(* IEC 61131-3 sources: Aqueous_Solutions/docs-authority/plc (part 3) *)

(* ---- PLC-HEAT.st ---- *)
(* AQS-CTL-004 X-CTL-04: control program source, generated by flow_graph/control/plc_programs.py *)
(* Basis: AQS-CTL-001 INSTRUMENT_INDEX.csv, AQS-CTL-002 control architecture, graph set-points. *)
(* PLC-HEAT: CPU single; IO counts AI 24 AO 0 DI 0 DO 0 (modules per AQS-CTL-002, 16-channel, 20 % spare) *)
PROGRAM PLC_HEAT_CTRL
VAR
  (* 100 ms cyclic task per AQS-CTL-002 *)
  DRY_COOLERPT-01_PV : REAL ;  (* no design pressure on the graph )
  DRY_COOLERTE-01_PV : REAL ;  (* band by service )
  Q1_APT-01_PV : REAL ;  (* no design pressure on the graph )
  Q1_ATE-01_PV : REAL ;  (* band by service )
  Q1_BPT-01_PV : REAL ;  (* no design pressure on the graph )
  Q1_BTE-01_PV : REAL ;  (* band by service )
  Q2_APT-01_PV : REAL ;  (* no design pressure on the graph )
  Q2_ATE-01_PV : REAL ;  (* band by service )
  Q2_BPT-01_PV : REAL ;  (* no design pressure on the graph )
  Q2_BTE-01_PV : REAL ;  (* band by service )
  Q3_APT-01_PV : REAL ;  (* no design pressure on the graph )
  Q3_ATE-01_PV : REAL ;  (* band by service )
  Q3_BPT-01_PV : REAL ;  (* no design pressure on the graph )
  Q3_BTE-01_PV : REAL ;  (* band by service )
  Q4_APT-01_PV : REAL ;  (* no design pressure on the graph )
  Q4_ATE-01_PV : REAL ;  (* band by service )
  Q4_BPT-01_PV : REAL ;  (* no design pressure on the graph )
  Q4_BTE-01_PV : REAL ;  (* band by service )
  ADS_CHILLTE-01_PV : REAL ;  (* drive water in: IA-Q4-ADS 5.0 kW Q4 65 C )
  ADS_CHILLTE-02_PV : REAL ;  (* chilled water out: IA-ADS-CHW 2.25 kW at 12 C )
  MAU_HXTE-01_PV : REAL ;  (* Q4 coil: IA-Q4-MAU 12 kW Q4 water 65/45 C (winter design) )
  Q4_BUSTE-01_PV : REAL ;  (* Q4 hot-water bus supply (IA-Q4-ADS/IA-Q4-MAU 65 C design) )
  Q4_BUSPT-01_PV : REAL ;  (* hot-water bus; no design pressure on the graph )
  RAD_PANELTE-01_PV : REAL ;  (* radiator loop outlet temperature watch; rejection performance against the A-M-39 )
END_VAR

  (* PRESSURE monitoring block - indication, no set-point invented )
  FB_AI_DRY_COOLERPT-01( PV := DRY_COOLERPT-01_PV );
  DRY_COOLERPT-01_ALARM_HI := 9.0 ;  (* 90 % of span, registered LSH convention )

  (* TEMPERATURE monitoring block - indication, no set-point invented )
  FB_AI_DRY_COOLERTE-01( PV := DRY_COOLERTE-01_PV );
  DRY_COOLERTE-01_ALARM_HI := 135.0 ;  (* 90 % of span, registered LSH convention )

  (* PRESSURE monitoring block - indication, no set-point invented )
  FB_AI_Q1_APT-01( PV := Q1_APT-01_PV );
  Q1_APT-01_ALARM_HI := 9.0 ;  (* 90 % of span, registered LSH convention )

  (* TEMPERATURE monitoring block - indication, no set-point invented )
  FB_AI_Q1_ATE-01( PV := Q1_ATE-01_PV );
  Q1_ATE-01_ALARM_HI := 135.0 ;  (* 90 % of span, registered LSH convention )

  (* PRESSURE monitoring block - indication, no set-point invented )
  FB_AI_Q1_BPT-01( PV := Q1_BPT-01_PV );
  Q1_BPT-01_ALARM_HI := 9.0 ;  (* 90 % of span, registered LSH convention )

  (* TEMPERATURE monitoring block - indication, no set-point invented )
  FB_AI_Q1_BTE-01( PV := Q1_BTE-01_PV );
  Q1_BTE-01_ALARM_HI := 135.0 ;  (* 90 % of span, registered LSH convention )

  (* PRESSURE monitoring block - indication, no set-point invented )
  FB_AI_Q2_APT-01( PV := Q2_APT-01_PV );
  Q2_APT-01_ALARM_HI := 9.0 ;  (* 90 % of span, registered LSH convention )

  (* TEMPERATURE monitoring block - indication, no set-point invented )
  FB_AI_Q2_ATE-01( PV := Q2_ATE-01_PV );
  Q2_ATE-01_ALARM_HI := 135.0 ;  (* 90 % of span, registered LSH convention )

  (* PRESSURE monitoring block - indication, no set-point invented )
  FB_AI_Q2_BPT-01( PV := Q2_BPT-01_PV );
  Q2_BPT-01_ALARM_HI := 9.0 ;  (* 90 % of span, registered LSH convention )

  (* TEMPERATURE monitoring block - indication, no set-point invented )
  FB_AI_Q2_BTE-01( PV := Q2_BTE-01_PV );
  Q2_BTE-01_ALARM_HI := 135.0 ;  (* 90 % of span, registered LSH convention )

  (* PRESSURE monitoring block - indication, no set-point invented )
  FB_AI_Q3_APT-01( PV := Q3_APT-01_PV );
  Q3_APT-01_ALARM_HI := 9.0 ;  (* 90 % of span, registered LSH convention )

  (* TEMPERATURE monitoring block - indication, no set-point invented )
  FB_AI_Q3_ATE-01( PV := Q3_ATE-01_PV );
  Q3_ATE-01_ALARM_HI := 135.0 ;  (* 90 % of span, registered LSH convention )

  (* PRESSURE monitoring block - indication, no set-point invented )
  FB_AI_Q3_BPT-01( PV := Q3_BPT-01_PV );
  Q3_BPT-01_ALARM_HI := 9.0 ;  (* 90 % of span, registered LSH convention )

  (* TEMPERATURE monitoring block - indication, no set-point invented )
  FB_AI_Q3_BTE-01( PV := Q3_BTE-01_PV );
  Q3_BTE-01_ALARM_HI := 135.0 ;  (* 90 % of span, registered LSH convention )

  (* PRESSURE monitoring block - indication, no set-point invented )
  FB_AI_Q4_APT-01( PV := Q4_APT-01_PV );
  Q4_APT-01_ALARM_HI := 9.0 ;  (* 90 % of span, registered LSH convention )

  (* TEMPERATURE monitoring block - indication, no set-point invented )
  FB_AI_Q4_ATE-01( PV := Q4_ATE-01_PV );
  Q4_ATE-01_ALARM_HI := 135.0 ;  (* 90 % of span, registered LSH convention )

  (* PRESSURE monitoring block - indication, no set-point invented )
  FB_AI_Q4_BPT-01( PV := Q4_BPT-01_PV );
  Q4_BPT-01_ALARM_HI := 9.0 ;  (* 90 % of span, registered LSH convention )

  (* TEMPERATURE monitoring block - indication, no set-point invented )
  FB_AI_Q4_BTE-01( PV := Q4_BTE-01_PV );
  Q4_BTE-01_ALARM_HI := 135.0 ;  (* 90 % of span, registered LSH convention )

  (* TEMPERATURE monitoring block - indication, no set-point invented )
  FB_AI_ADS_CHILLTE-01( PV := ADS_CHILLTE-01_PV );
  ADS_CHILLTE-01_ALARM_HI := 90.0 ;  (* 90 % of span, registered LSH convention )

  (* TEMPERATURE monitoring block - indication, no set-point invented )
  FB_AI_ADS_CHILLTE-02( PV := ADS_CHILLTE-02_PV );
  ADS_CHILLTE-02_ALARM_HI := 36.0 ;  (* 90 % of span, registered LSH convention )

  (* TEMPERATURE monitoring block - indication, no set-point invented )
  FB_AI_MAU_HXTE-01( PV := MAU_HXTE-01_PV );
  MAU_HXTE-01_ALARM_HI := 90.0 ;  (* 90 % of span, registered LSH convention )

  (* TEMPERATURE monitoring block - indication, no set-point invented )
  FB_AI_Q4_BUSTE-01( PV := Q4_BUSTE-01_PV );
  Q4_BUSTE-01_ALARM_HI := 90.0 ;  (* 90 % of span, registered LSH convention )

  (* PRESSURE monitoring block - indication, no set-point invented )
  FB_AI_Q4_BUSPT-01( PV := Q4_BUSPT-01_PV );
  Q4_BUSPT-01_ALARM_HI := 9.0 ;  (* 90 % of span, registered LSH convention )

  (* TEMPERATURE monitoring block - indication, no set-point invented )
  FB_AI_RAD_PANELTE-01( PV := RAD_PANELTE-01_PV );
  RAD_PANELTE-01_ALARM_HI := 135.0 ;  (* 90 % of span, registered LSH convention )

END_PROGRAM

(* ---- PLC-MEOH.st ---- *)
(* AQS-CTL-004 X-CTL-04: control program source, generated by flow_graph/control/plc_programs.py *)
(* Basis: AQS-CTL-001 INSTRUMENT_INDEX.csv, AQS-CTL-002 control architecture, graph set-points. *)
(* PLC-MEOH: CPU single; IO counts AI 33 AO 0 DI 51 DO 12 (modules per AQS-CTL-002, 16-channel, 20 % spare) *)
PROGRAM PLC_MEOH_CTRL
VAR
  (* 100 ms cyclic task per AQS-CTL-002 *)
  MET_SYNFT-01_PV : REAL ;  (* DL_MET_TO_FEED normal 0.00 L/h )
  MET_SYNPT-01_PV : REAL ;  (* no design pressure on the graph )
  MET_SYNTE-01_PV : REAL ;  (* band by service )
  MEOH_FERMFT-01_PV : REAL ;  (* S77 normal 0.00 L/h )
  MEOH_FERMPT-01_PV : REAL ;  (* no design pressure on the graph )
  MEOH_FERMTE-01_PV : REAL ;  (* design T 35 C )
  MEOH_FCFT-01_PV : REAL ;  (* S81 normal 0.30 L/h )
  MEOH_FCFT-02_PV : REAL ;  (* S82 normal 0.36 L/h )
  MEOH_FCFT-03_PV : REAL ;  (* IA-FC-EXH normal 0.00 L/h )
  MEOH_FCLT-01_PV : REAL ;  (* A-M-182 liquid height )
  MEOH_FCPT-01_PV : REAL ;  (* no design pressure on the graph )
  MEOH_FCTE-01_PV : REAL ;  (* band by service )
  MEOH_SYNTHFT-01_PV : REAL ;  (* IA-ESS-MEOH-CHG normal 0.00 L/h )
  MEOH_SYNTHFT-02_PV : REAL ;  (* S75 normal 1.47 L/h )
  MEOH_SYNTHFT-03_PV : REAL ;  (* MEOH_TO_OLEFIN normal 0.00 L/h )
  MEOH_SYNTHFT-04_PV : REAL ;  (* IA-MEOH-H2O normal 0.82 L/h )
  MEOH_SYNTHFT-05_PV : REAL ;  (* IA-MEOH-CH3SH normal 0.00 L/h )
  MEOH_SYNTHPT-01_PV : REAL ;  (* no design pressure on the graph )
  MEOH_SYNTHTE-01_PV : REAL ;  (* design T 250 C )
  MEOH_CONDLT-01_PV : REAL ;  (* A-M-182 liquid height )
  MEOH_CONDPT-01_PV : REAL ;  (* no design pressure on the graph )
  MEOH_CONDTE-01_PV : REAL ;  (* band by service )
  MEOH_TANKFT-01_PV : REAL ;  (* S76 normal 0.21 L/h )
  MEOH_TANKFT-02_PV : REAL ;  (* IA-MEOH-REST normal 0.05 L/h )
  MEOH_TANKFT-03_PV : REAL ;  (* IA-MEOH-PROD normal 1.19 L/h )
  MEOH_TANKFT-04_PV : REAL ;  (* MEOH_TO_VDF normal 0.01 L/h )
  MEOH_TANKFT-05_PV : REAL ;  (* MEOH_TO_TFE normal 0.00 L/h )
  MEOH_TANKLT-01_PV : REAL ;  (* A-M-182 liquid height )
  MEOH_TANKPT-01_PV : REAL ;  (* no design pressure on the graph )
  MEOH_TANKTE-01_PV : REAL ;  (* band by service )
  MET_SYNTIR-01_PV : REAL ;  (* the Strecker step is temperature-sensitive: the hydrolysis runs at 100-150 C (X- )
  MET_SYNFIT-01_PV : REAL ;  (* the precursor metering: CH3SH, acrolein and NH3 are each fed at the gram/h class )
  MEOH_SYNTHTE-90 : BOOL ;  (* SIF watch input, routed to the safety CPU pair (AQS-CTL-003) *)
END_VAR

  (* FLOW control loop - set-point from the graph basis *)
  MET_SYNFT-01_SP := 0.0 ;  (* graph basis: DL_MET_TO_FEED normal 0.00 L/h )
  FB_PI_MET_SYNFT-01( PV := MET_SYNFT-01_PV, SP := MET_SYNFT-01_SP );  (* PI per AQS-CTL-002; GAIN/KI entered at commissioning from the step test (AQS-COM-001 sec. 3), anti-windup clamp per this FB *)
  MET_SYNFT-01_ALARM_HI := 0.0 ;  (* expected-zero state: any positive PV alarms )

  (* PRESSURE monitoring block - indication, no set-point invented )
  FB_AI_MET_SYNPT-01( PV := MET_SYNPT-01_PV );
  MET_SYNPT-01_ALARM_HI := 9.0 ;  (* 90 % of span, registered LSH convention )

  (* TEMPERATURE monitoring block - indication, no set-point invented )
  FB_AI_MET_SYNTE-01( PV := MET_SYNTE-01_PV );
  MET_SYNTE-01_ALARM_HI := 135.0 ;  (* 90 % of span, registered LSH convention )

  (* FLOW control loop - set-point from the graph basis *)
  MEOH_FERMFT-01_SP := 0.0 ;  (* graph basis: S77 normal 0.00 L/h )
  FB_PI_MEOH_FERMFT-01( PV := MEOH_FERMFT-01_PV, SP := MEOH_FERMFT-01_SP );  (* PI per AQS-CTL-002; GAIN/KI entered at commissioning from the step test (AQS-COM-001 sec. 3), anti-windup clamp per this FB *)
  MEOH_FERMFT-01_ALARM_HI := 0.0 ;  (* expected-zero state: any positive PV alarms )

  (* PRESSURE monitoring block - indication, no set-point invented )
  FB_AI_MEOH_FERMPT-01( PV := MEOH_FERMPT-01_PV );
  MEOH_FERMPT-01_ALARM_HI := 9.0 ;  (* 90 % of span, registered LSH convention )

  (* TEMPERATURE control loop - set-point from the graph basis *)
  MEOH_FERMTE-01_SP := 35.0 ;  (* graph basis: design T 35 C )
  FB_PI_MEOH_FERMTE-01( PV := MEOH_FERMTE-01_PV, SP := MEOH_FERMTE-01_SP );  (* PI per AQS-CTL-002; GAIN/KI entered at commissioning from the step test (AQS-COM-001 sec. 3), anti-windup clamp per this FB *)
  MEOH_FERMTE-01_ALARM_HI := 38.5 ;  (* SP x 1.1 margin, A-M-188 margin class *)
  MEOH_FERMTE-01_ALARM_LO := 31.5 ;

  (* FLOW control loop - set-point from the graph basis *)
  MEOH_FCFT-01_SP := 0.3 ;  (* graph basis: S81 normal 0.30 L/h )
  FB_PI_MEOH_FCFT-01( PV := MEOH_FCFT-01_PV, SP := MEOH_FCFT-01_SP );  (* PI per AQS-CTL-002; GAIN/KI entered at commissioning from the step test (AQS-COM-001 sec. 3), anti-windup clamp per this FB *)
  MEOH_FCFT-01_ALARM_HI := 0.33 ;  (* SP x 1.1 margin, A-M-188 margin class *)
  MEOH_FCFT-01_ALARM_LO := 0.27 ;

  (* FLOW control loop - set-point from the graph basis *)
  MEOH_FCFT-02_SP := 0.36 ;  (* graph basis: S82 normal 0.36 L/h )
  FB_PI_MEOH_FCFT-02( PV := MEOH_FCFT-02_PV, SP := MEOH_FCFT-02_SP );  (* PI per AQS-CTL-002; GAIN/KI entered at commissioning from the step test (AQS-COM-001 sec. 3), anti-windup clamp per this FB *)
  MEOH_FCFT-02_ALARM_HI := 0.396 ;  (* SP x 1.1 margin, A-M-188 margin class *)
  MEOH_FCFT-02_ALARM_LO := 0.324 ;

  (* FLOW control loop - set-point from the graph basis *)
  MEOH_FCFT-03_SP := 0.0 ;  (* graph basis: IA-FC-EXH normal 0.00 L/h )
  FB_PI_MEOH_FCFT-03( PV := MEOH_FCFT-03_PV, SP := MEOH_FCFT-03_SP );  (* PI per AQS-CTL-002; GAIN/KI entered at commissioning from the step test (AQS-COM-001 sec. 3), anti-windup clamp per this FB *)
  MEOH_FCFT-03_ALARM_HI := 0.0 ;  (* expected-zero state: any positive PV alarms )

  (* LEVEL monitoring block - indication, no set-point invented )
  FB_AI_MEOH_FCLT-01( PV := MEOH_FCLT-01_PV );
  MEOH_FCLT-01_ALARM_HI := 90.0 ;  (* 90 % of span, registered LSH convention )

  (* PRESSURE monitoring block - indication, no set-point invented )
  FB_AI_MEOH_FCPT-01( PV := MEOH_FCPT-01_PV );
  MEOH_FCPT-01_ALARM_HI := 9.0 ;  (* 90 % of span, registered LSH convention )

  (* TEMPERATURE monitoring block - indication, no set-point invented )
  FB_AI_MEOH_FCTE-01( PV := MEOH_FCTE-01_PV );
  MEOH_FCTE-01_ALARM_HI := 135.0 ;  (* 90 % of span, registered LSH convention )

  (* FLOW control loop - set-point from the graph basis *)
  MEOH_SYNTHFT-01_SP := 0.0 ;  (* graph basis: IA-ESS-MEOH-CHG normal 0.00 L/h )
  FB_PI_MEOH_SYNTHFT-01( PV := MEOH_SYNTHFT-01_PV, SP := MEOH_SYNTHFT-01_SP );  (* PI per AQS-CTL-002; GAIN/KI entered at commissioning from the step test (AQS-COM-001 sec. 3), anti-windup clamp per this FB *)
  MEOH_SYNTHFT-01_ALARM_HI := 0.0 ;  (* expected-zero state: any positive PV alarms )

  (* FLOW control loop - set-point from the graph basis *)
  MEOH_SYNTHFT-02_SP := 1.47 ;  (* graph basis: S75 normal 1.47 L/h )
  FB_PI_MEOH_SYNTHFT-02( PV := MEOH_SYNTHFT-02_PV, SP := MEOH_SYNTHFT-02_SP );  (* PI per AQS-CTL-002; GAIN/KI entered at commissioning from the step test (AQS-COM-001 sec. 3), anti-windup clamp per this FB *)
  MEOH_SYNTHFT-02_ALARM_HI := 1.617 ;  (* SP x 1.1 margin, A-M-188 margin class *)
  MEOH_SYNTHFT-02_ALARM_LO := 1.323 ;

  (* FLOW control loop - set-point from the graph basis *)
  MEOH_SYNTHFT-03_SP := 0.0 ;  (* graph basis: MEOH_TO_OLEFIN normal 0.00 L/h )
  FB_PI_MEOH_SYNTHFT-03( PV := MEOH_SYNTHFT-03_PV, SP := MEOH_SYNTHFT-03_SP );  (* PI per AQS-CTL-002; GAIN/KI entered at commissioning from the step test (AQS-COM-001 sec. 3), anti-windup clamp per this FB *)
  MEOH_SYNTHFT-03_ALARM_HI := 0.0 ;  (* expected-zero state: any positive PV alarms )

  (* FLOW control loop - set-point from the graph basis *)
  MEOH_SYNTHFT-04_SP := 0.82 ;  (* graph basis: IA-MEOH-H2O normal 0.82 L/h )
  FB_PI_MEOH_SYNTHFT-04( PV := MEOH_SYNTHFT-04_PV, SP := MEOH_SYNTHFT-04_SP );  (* PI per AQS-CTL-002; GAIN/KI entered at commissioning from the step test (AQS-COM-001 sec. 3), anti-windup clamp per this FB *)
  MEOH_SYNTHFT-04_ALARM_HI := 0.902 ;  (* SP x 1.1 margin, A-M-188 margin class *)
  MEOH_SYNTHFT-04_ALARM_LO := 0.738 ;

  (* FLOW control loop - set-point from the graph basis *)
  MEOH_SYNTHFT-05_SP := 0.0 ;  (* graph basis: IA-MEOH-CH3SH normal 0.00 L/h )
  FB_PI_MEOH_SYNTHFT-05( PV := MEOH_SYNTHFT-05_PV, SP := MEOH_SYNTHFT-05_SP );  (* PI per AQS-CTL-002; GAIN/KI entered at commissioning from the step test (AQS-COM-001 sec. 3), anti-windup clamp per this FB *)
  MEOH_SYNTHFT-05_ALARM_HI := 0.0 ;  (* expected-zero state: any positive PV alarms )

  (* PRESSURE monitoring block - indication, no set-point invented )
  FB_AI_MEOH_SYNTHPT-01( PV := MEOH_SYNTHPT-01_PV );
  MEOH_SYNTHPT-01_ALARM_HI := 9.0 ;  (* 90 % of span, registered LSH convention )

  (* TEMPERATURE control loop - set-point from the graph basis *)
  MEOH_SYNTHTE-01_SP := 250.0 ;  (* graph basis: design T 250 C )
  FB_PI_MEOH_SYNTHTE-01( PV := MEOH_SYNTHTE-01_PV, SP := MEOH_SYNTHTE-01_SP );  (* PI per AQS-CTL-002; GAIN/KI entered at commissioning from the step test (AQS-COM-001 sec. 3), anti-windup clamp per this FB *)
  MEOH_SYNTHTE-01_ALARM_HI := 275.0 ;  (* SP x 1.1 margin, A-M-188 margin class *)
  MEOH_SYNTHTE-01_ALARM_LO := 225.0 ;

  (* LEVEL monitoring block - indication, no set-point invented )
  FB_AI_MEOH_CONDLT-01( PV := MEOH_CONDLT-01_PV );
  MEOH_CONDLT-01_ALARM_HI := 90.0 ;  (* 90 % of span, registered LSH convention )

  (* PRESSURE monitoring block - indication, no set-point invented )
  FB_AI_MEOH_CONDPT-01( PV := MEOH_CONDPT-01_PV );
  MEOH_CONDPT-01_ALARM_HI := 9.0 ;  (* 90 % of span, registered LSH convention )

  (* TEMPERATURE monitoring block - indication, no set-point invented )
  FB_AI_MEOH_CONDTE-01( PV := MEOH_CONDTE-01_PV );
  MEOH_CONDTE-01_ALARM_HI := 135.0 ;  (* 90 % of span, registered LSH convention )

  (* FLOW control loop - set-point from the graph basis *)
  MEOH_TANKFT-01_SP := 0.21 ;  (* graph basis: S76 normal 0.21 L/h )
  FB_PI_MEOH_TANKFT-01( PV := MEOH_TANKFT-01_PV, SP := MEOH_TANKFT-01_SP );  (* PI per AQS-CTL-002; GAIN/KI entered at commissioning from the step test (AQS-COM-001 sec. 3), anti-windup clamp per this FB *)
  MEOH_TANKFT-01_ALARM_HI := 0.231 ;  (* SP x 1.1 margin, A-M-188 margin class *)
  MEOH_TANKFT-01_ALARM_LO := 0.189 ;

  (* FLOW control loop - set-point from the graph basis *)
  MEOH_TANKFT-02_SP := 0.05 ;  (* graph basis: IA-MEOH-REST normal 0.05 L/h )
  FB_PI_MEOH_TANKFT-02( PV := MEOH_TANKFT-02_PV, SP := MEOH_TANKFT-02_SP );  (* PI per AQS-CTL-002; GAIN/KI entered at commissioning from the step test (AQS-COM-001 sec. 3), anti-windup clamp per this FB *)
  MEOH_TANKFT-02_ALARM_HI := 0.05500000000000001 ;  (* SP x 1.1 margin, A-M-188 margin class *)
  MEOH_TANKFT-02_ALARM_LO := 0.045000000000000005 ;

  (* FLOW control loop - set-point from the graph basis *)
  MEOH_TANKFT-03_SP := 1.19 ;  (* graph basis: IA-MEOH-PROD normal 1.19 L/h )
  FB_PI_MEOH_TANKFT-03( PV := MEOH_TANKFT-03_PV, SP := MEOH_TANKFT-03_SP );  (* PI per AQS-CTL-002; GAIN/KI entered at commissioning from the step test (AQS-COM-001 sec. 3), anti-windup clamp per this FB *)
  MEOH_TANKFT-03_ALARM_HI := 1.309 ;  (* SP x 1.1 margin, A-M-188 margin class *)
  MEOH_TANKFT-03_ALARM_LO := 1.071 ;

  (* FLOW control loop - set-point from the graph basis *)
  MEOH_TANKFT-04_SP := 0.01 ;  (* graph basis: MEOH_TO_VDF normal 0.01 L/h )
  FB_PI_MEOH_TANKFT-04( PV := MEOH_TANKFT-04_PV, SP := MEOH_TANKFT-04_SP );  (* PI per AQS-CTL-002; GAIN/KI entered at commissioning from the step test (AQS-COM-001 sec. 3), anti-windup clamp per this FB *)
  MEOH_TANKFT-04_ALARM_HI := 0.011000000000000001 ;  (* SP x 1.1 margin, A-M-188 margin class *)
  MEOH_TANKFT-04_ALARM_LO := 0.009000000000000001 ;

  (* FLOW control loop - set-point from the graph basis *)
  MEOH_TANKFT-05_SP := 0.0 ;  (* graph basis: MEOH_TO_TFE normal 0.00 L/h )
  FB_PI_MEOH_TANKFT-05( PV := MEOH_TANKFT-05_PV, SP := MEOH_TANKFT-05_SP );  (* PI per AQS-CTL-002; GAIN/KI entered at commissioning from the step test (AQS-COM-001 sec. 3), anti-windup clamp per this FB *)
  MEOH_TANKFT-05_ALARM_HI := 0.0 ;  (* expected-zero state: any positive PV alarms )

  (* LEVEL monitoring block - indication, no set-point invented )
  FB_AI_MEOH_TANKLT-01( PV := MEOH_TANKLT-01_PV );
  MEOH_TANKLT-01_ALARM_HI := 90.0 ;  (* 90 % of span, registered LSH convention )

  (* PRESSURE monitoring block - indication, no set-point invented )
  FB_AI_MEOH_TANKPT-01( PV := MEOH_TANKPT-01_PV );
  MEOH_TANKPT-01_ALARM_HI := 9.0 ;  (* 90 % of span, registered LSH convention )

  (* TEMPERATURE monitoring block - indication, no set-point invented )
  FB_AI_MEOH_TANKTE-01( PV := MEOH_TANKTE-01_PV );
  MEOH_TANKTE-01_ALARM_HI := 135.0 ;  (* 90 % of span, registered LSH convention )

  (* TEMPERATURE monitoring block - indication, no set-point invented )
  FB_AI_MET_SYNTIR-01( PV := MET_SYNTIR-01_PV );
  MET_SYNTIR-01_ALARM_HI := 180.0 ;  (* 90 % of span, registered LSH convention )

  (* FLOW monitoring block - indication, no set-point invented )
  FB_AI_MET_SYNFIT-01( PV := MET_SYNFIT-01_PV );
  MET_SYNFIT-01_ALARM_HI := 45.0 ;  (* 90 % of span, registered LSH convention )

  (* SIF watch passthrough, no action in the basic program )
  SIF_WATCH_MEOH_SYNTHTE-90 := MEOH_SYNTHTE-90 ;  (* to safety CPU pair, AQS-CTL-003 )

END_PROGRAM

(* ---- PLC-MFG.st ---- *)
(* AQS-CTL-004 X-CTL-04: control program source, generated by flow_graph/control/plc_programs.py *)
(* Basis: AQS-CTL-001 INSTRUMENT_INDEX.csv, AQS-CTL-002 control architecture, graph set-points. *)
(* PLC-MFG: CPU single; IO counts AI 32 AO 9 DI 42 DO 5 (modules per AQS-CTL-002, 16-channel, 20 % spare) *)
PROGRAM PLC_MFG_CTRL
VAR
  (* 100 ms cyclic task per AQS-CTL-002 *)
  COLD_MILLPT-01_PV : REAL ;  (* no design pressure on the graph )
  COLD_MILLTE-01_PV : REAL ;  (* band by service )
  GAS_ATOMIZERPT-01_PV : REAL ;  (* no design pressure on the graph )
  GAS_ATOMIZERTE-01_PV : REAL ;  (* band by service )
  MET_MELTFT-01_PV : REAL ;  (* S57 normal 0.15 L/h )
  MET_MELTPT-01_PV : REAL ;  (* no design pressure on the graph )
  MET_MELTTE-01_PV : REAL ;  (* band by service )
  MFG_SHOPFT-01_PV : REAL ;  (* TEXTILE_HAB normal 0.00 L/h )
  MFG_SHOPLT-01_PV : REAL ;  (* A-M-182 liquid height )
  MFG_SHOPPT-01_PV : REAL ;  (* no design pressure on the graph )
  MFG_SHOPTE-01_PV : REAL ;  (* band by service )
  WIRE_DRAWPT-01_PV : REAL ;  (* no design pressure on the graph )
  WIRE_DRAWTE-01_PV : REAL ;  (* band by service )
  MET_AHUPT-01_PV : REAL ;  (* no design pressure on the graph )
  MET_AHUTE-01_PV : REAL ;  (* band by service )
  ELECTRODE_COATPT-01_PV : REAL ;  (* no design pressure on the graph )
  ELECTRODE_COATTE-01_PV : REAL ;  (* band by service )
  BLOW_MOLDPT-01_PV : REAL ;  (* no design pressure on the graph )
  BLOW_MOLDTE-01_PV : REAL ;  (* band by service )
  MET_HX_Q4PT-01_PV : REAL ;  (* no design pressure on the graph )
  MET_HX_Q4TE-01_PV : REAL ;  (* band by service )
  REE_RECOVERPT-01_PV : REAL ;  (* no design pressure on the graph )
  REE_RECOVERTE-01_PV : REAL ;  (* band by service )
  MET_SCRUBFT-01_PV : REAL ;  (* S72 normal 0.10 L/h )
  MET_SCRUBFT-02_PV : REAL ;  (* S72B normal 0.00 L/h )
  MET_SCRUBFT-03_PV : REAL ;  (* IA-MET-AIR-RET normal 2983.40 L/h )
  MET_SCRUBLT-01_PV : REAL ;  (* A-M-182 liquid height )
  MET_SCRUBPT-01_PV : REAL ;  (* no design pressure on the graph )
  MET_SCRUBTE-01_PV : REAL ;  (* band by service )
  REE_RECOVERTIR-01_PV : REAL ;  (* campaign temperature control: leach 55 C, demag > 320 C (Nd2Fe14B Curie), calcin )
  REE_RECOVERSIT-01_PV : REAL ;  (* pH fronts the two precipitations: Fe(OH)3 sweep at pH 3-3.5, RE oxalate at pH 1- )
  MET_MELTTE-90 : BOOL ;  (* SIF watch input, routed to the safety CPU pair (AQS-CTL-003) *)
END_VAR

  (* PRESSURE monitoring block - indication, no set-point invented )
  FB_AI_COLD_MILLPT-01( PV := COLD_MILLPT-01_PV );
  COLD_MILLPT-01_ALARM_HI := 9.0 ;  (* 90 % of span, registered LSH convention )

  (* TEMPERATURE monitoring block - indication, no set-point invented )
  FB_AI_COLD_MILLTE-01( PV := COLD_MILLTE-01_PV );
  COLD_MILLTE-01_ALARM_HI := 135.0 ;  (* 90 % of span, registered LSH convention )

  (* PRESSURE monitoring block - indication, no set-point invented )
  FB_AI_GAS_ATOMIZERPT-01( PV := GAS_ATOMIZERPT-01_PV );
  GAS_ATOMIZERPT-01_ALARM_HI := 9.0 ;  (* 90 % of span, registered LSH convention )

  (* TEMPERATURE monitoring block - indication, no set-point invented )
  FB_AI_GAS_ATOMIZERTE-01( PV := GAS_ATOMIZERTE-01_PV );
  GAS_ATOMIZERTE-01_ALARM_HI := 135.0 ;  (* 90 % of span, registered LSH convention )

  (* FLOW control loop - set-point from the graph basis *)
  MET_MELTFT-01_SP := 0.15 ;  (* graph basis: S57 normal 0.15 L/h )
  FB_PI_MET_MELTFT-01( PV := MET_MELTFT-01_PV, SP := MET_MELTFT-01_SP );  (* PI per AQS-CTL-002; GAIN/KI entered at commissioning from the step test (AQS-COM-001 sec. 3), anti-windup clamp per this FB *)
  MET_MELTFT-01_ALARM_HI := 0.165 ;  (* SP x 1.1 margin, A-M-188 margin class *)
  MET_MELTFT-01_ALARM_LO := 0.135 ;

  (* PRESSURE monitoring block - indication, no set-point invented )
  FB_AI_MET_MELTPT-01( PV := MET_MELTPT-01_PV );
  MET_MELTPT-01_ALARM_HI := 9.0 ;  (* 90 % of span, registered LSH convention )

  (* TEMPERATURE monitoring block - indication, no set-point invented )
  FB_AI_MET_MELTTE-01( PV := MET_MELTTE-01_PV );
  MET_MELTTE-01_ALARM_HI := 540.0 ;  (* 90 % of span, registered LSH convention )

  (* FLOW control loop - set-point from the graph basis *)
  MFG_SHOPFT-01_SP := 0.0 ;  (* graph basis: TEXTILE_HAB normal 0.00 L/h )
  FB_PI_MFG_SHOPFT-01( PV := MFG_SHOPFT-01_PV, SP := MFG_SHOPFT-01_SP );  (* PI per AQS-CTL-002; GAIN/KI entered at commissioning from the step test (AQS-COM-001 sec. 3), anti-windup clamp per this FB *)
  MFG_SHOPFT-01_ALARM_HI := 0.0 ;  (* expected-zero state: any positive PV alarms )

  (* LEVEL monitoring block - indication, no set-point invented )
  FB_AI_MFG_SHOPLT-01( PV := MFG_SHOPLT-01_PV );
  MFG_SHOPLT-01_ALARM_HI := 90.0 ;  (* 90 % of span, registered LSH convention )

  (* PRESSURE monitoring block - indication, no set-point invented )
  FB_AI_MFG_SHOPPT-01( PV := MFG_SHOPPT-01_PV );
  MFG_SHOPPT-01_ALARM_HI := 9.0 ;  (* 90 % of span, registered LSH convention )

  (* TEMPERATURE monitoring block - indication, no set-point invented )
  FB_AI_MFG_SHOPTE-01( PV := MFG_SHOPTE-01_PV );
  MFG_SHOPTE-01_ALARM_HI := 135.0 ;  (* 90 % of span, registered LSH convention )

  (* PRESSURE monitoring block - indication, no set-point invented )
  FB_AI_WIRE_DRAWPT-01( PV := WIRE_DRAWPT-01_PV );
  WIRE_DRAWPT-01_ALARM_HI := 9.0 ;  (* 90 % of span, registered LSH convention )

  (* TEMPERATURE monitoring block - indication, no set-point invented )
  FB_AI_WIRE_DRAWTE-01( PV := WIRE_DRAWTE-01_PV );
  WIRE_DRAWTE-01_ALARM_HI := 135.0 ;  (* 90 % of span, registered LSH convention )

  (* PRESSURE monitoring block - indication, no set-point invented )
  FB_AI_MET_AHUPT-01( PV := MET_AHUPT-01_PV );
  MET_AHUPT-01_ALARM_HI := 9.0 ;  (* 90 % of span, registered LSH convention )

  (* TEMPERATURE monitoring block - indication, no set-point invented )
  FB_AI_MET_AHUTE-01( PV := MET_AHUTE-01_PV );
  MET_AHUTE-01_ALARM_HI := 135.0 ;  (* 90 % of span, registered LSH convention )

  (* PRESSURE monitoring block - indication, no set-point invented )
  FB_AI_ELECTRODE_COATPT-01( PV := ELECTRODE_COATPT-01_PV );
  ELECTRODE_COATPT-01_ALARM_HI := 9.0 ;  (* 90 % of span, registered LSH convention )

  (* TEMPERATURE monitoring block - indication, no set-point invented )
  FB_AI_ELECTRODE_COATTE-01( PV := ELECTRODE_COATTE-01_PV );
  ELECTRODE_COATTE-01_ALARM_HI := 135.0 ;  (* 90 % of span, registered LSH convention )

  (* PRESSURE monitoring block - indication, no set-point invented )
  FB_AI_BLOW_MOLDPT-01( PV := BLOW_MOLDPT-01_PV );
  BLOW_MOLDPT-01_ALARM_HI := 9.0 ;  (* 90 % of span, registered LSH convention )

  (* TEMPERATURE monitoring block - indication, no set-point invented )
  FB_AI_BLOW_MOLDTE-01( PV := BLOW_MOLDTE-01_PV );
  BLOW_MOLDTE-01_ALARM_HI := 135.0 ;  (* 90 % of span, registered LSH convention )

  (* PRESSURE monitoring block - indication, no set-point invented )
  FB_AI_MET_HX_Q4PT-01( PV := MET_HX_Q4PT-01_PV );
  MET_HX_Q4PT-01_ALARM_HI := 9.0 ;  (* 90 % of span, registered LSH convention )

  (* TEMPERATURE monitoring block - indication, no set-point invented )
  FB_AI_MET_HX_Q4TE-01( PV := MET_HX_Q4TE-01_PV );
  MET_HX_Q4TE-01_ALARM_HI := 135.0 ;  (* 90 % of span, registered LSH convention )

  (* PRESSURE monitoring block - indication, no set-point invented )
  FB_AI_REE_RECOVERPT-01( PV := REE_RECOVERPT-01_PV );
  REE_RECOVERPT-01_ALARM_HI := 9.0 ;  (* 90 % of span, registered LSH convention )

  (* TEMPERATURE monitoring block - indication, no set-point invented )
  FB_AI_REE_RECOVERTE-01( PV := REE_RECOVERTE-01_PV );
  REE_RECOVERTE-01_ALARM_HI := 135.0 ;  (* 90 % of span, registered LSH convention )

  (* FLOW control loop - set-point from the graph basis *)
  MET_SCRUBFT-01_SP := 0.1 ;  (* graph basis: S72 normal 0.10 L/h )
  FB_PI_MET_SCRUBFT-01( PV := MET_SCRUBFT-01_PV, SP := MET_SCRUBFT-01_SP );  (* PI per AQS-CTL-002; GAIN/KI entered at commissioning from the step test (AQS-COM-001 sec. 3), anti-windup clamp per this FB *)
  MET_SCRUBFT-01_ALARM_HI := 0.11000000000000001 ;  (* SP x 1.1 margin, A-M-188 margin class *)
  MET_SCRUBFT-01_ALARM_LO := 0.09000000000000001 ;

  (* FLOW control loop - set-point from the graph basis *)
  MET_SCRUBFT-02_SP := 0.0 ;  (* graph basis: S72B normal 0.00 L/h )
  FB_PI_MET_SCRUBFT-02( PV := MET_SCRUBFT-02_PV, SP := MET_SCRUBFT-02_SP );  (* PI per AQS-CTL-002; GAIN/KI entered at commissioning from the step test (AQS-COM-001 sec. 3), anti-windup clamp per this FB *)
  MET_SCRUBFT-02_ALARM_HI := 0.0 ;  (* expected-zero state: any positive PV alarms )

  (* FLOW control loop - set-point from the graph basis *)
  MET_SCRUBFT-03_SP := 2983.4 ;  (* graph basis: IA-MET-AIR-RET normal 2983.40 L/h )
  FB_PI_MET_SCRUBFT-03( PV := MET_SCRUBFT-03_PV, SP := MET_SCRUBFT-03_SP );  (* PI per AQS-CTL-002; GAIN/KI entered at commissioning from the step test (AQS-COM-001 sec. 3), anti-windup clamp per this FB *)
  MET_SCRUBFT-03_ALARM_HI := 3281.7400000000002 ;  (* SP x 1.1 margin, A-M-188 margin class *)
  MET_SCRUBFT-03_ALARM_LO := 2685.06 ;

  (* LEVEL monitoring block - indication, no set-point invented )
  FB_AI_MET_SCRUBLT-01( PV := MET_SCRUBLT-01_PV );
  MET_SCRUBLT-01_ALARM_HI := 90.0 ;  (* 90 % of span, registered LSH convention )

  (* PRESSURE monitoring block - indication, no set-point invented )
  FB_AI_MET_SCRUBPT-01( PV := MET_SCRUBPT-01_PV );
  MET_SCRUBPT-01_ALARM_HI := 9.0 ;  (* 90 % of span, registered LSH convention )

  (* TEMPERATURE monitoring block - indication, no set-point invented )
  FB_AI_MET_SCRUBTE-01( PV := MET_SCRUBTE-01_PV );
  MET_SCRUBTE-01_ALARM_HI := 135.0 ;  (* 90 % of span, registered LSH convention )

  (* TEMPERATURE monitoring block - indication, no set-point invented )
  FB_AI_REE_RECOVERTIR-01( PV := REE_RECOVERTIR-01_PV );
  REE_RECOVERTIR-01_ALARM_HI := 900.0 ;  (* 90 % of span, registered LSH convention )

  (* PH monitoring block - indication, no set-point invented )
  FB_AI_REE_RECOVERSIT-01( PV := REE_RECOVERSIT-01_PV );
  REE_RECOVERSIT-01_ALARM_HI := 12.6 ;  (* 90 % of span, registered LSH convention )

  (* SIF watch passthrough, no action in the basic program )
  SIF_WATCH_MET_MELTTE-90 := MET_MELTTE-90 ;  (* to safety CPU pair, AQS-CTL-003 )

END_PROGRAM

(* ---- PLC-NUT.st ---- *)
(* AQS-CTL-004 X-CTL-04: control program source, generated by flow_graph/control/plc_programs.py *)
(* Basis: AQS-CTL-001 INSTRUMENT_INDEX.csv, AQS-CTL-002 control architecture, graph set-points. *)
(* PLC-NUT: CPU redundant pair; IO counts AI 9 AO 0 DI 11 DO 5 (modules per AQS-CTL-002, 16-channel, 20 % spare) *)
PROGRAM PLC_NUT_CTRL
VAR
  (* 100 ms cyclic task per AQS-CTL-002 *)
  NUTRIENT_DOSEFT-01_PV : REAL ;  (* S07 normal 0.10 L/h )
  NUTRIENT_DOSEFT-02_PV : REAL ;  (* NUT_TO_BED normal 0.00 L/h )
  NUTRIENT_DOSEFT-03_PV : REAL ;  (* IA-NUT-01 normal 0.58 L/h )
  NUTRIENT_DOSEFT-04_PV : REAL ;  (* IA-NUT-LEACH normal 3.43 L/h )
  NUTRIENT_DOSEFT-05_PV : REAL ;  (* IA-NUT-BED normal 1.31 L/h )
  NUTRIENT_DOSEFT-06_PV : REAL ;  (* IA-SIC-RET normal 0.02 L/h )
  NUTRIENT_DOSELT-01_PV : REAL ;  (* A-M-182 liquid height )
  NUTRIENT_DOSEPT-01_PV : REAL ;  (* no design pressure on the graph )
  NUTRIENT_DOSETE-01_PV : REAL ;  (* band by service )
END_VAR

  (* FLOW control loop - set-point from the graph basis *)
  NUTRIENT_DOSEFT-01_SP := 0.1 ;  (* graph basis: S07 normal 0.10 L/h )
  FB_PI_NUTRIENT_DOSEFT-01( PV := NUTRIENT_DOSEFT-01_PV, SP := NUTRIENT_DOSEFT-01_SP );  (* PI per AQS-CTL-002; GAIN/KI entered at commissioning from the step test (AQS-COM-001 sec. 3), anti-windup clamp per this FB *)
  NUTRIENT_DOSEFT-01_ALARM_HI := 0.11000000000000001 ;  (* SP x 1.1 margin, A-M-188 margin class *)
  NUTRIENT_DOSEFT-01_ALARM_LO := 0.09000000000000001 ;

  (* FLOW control loop - set-point from the graph basis *)
  NUTRIENT_DOSEFT-02_SP := 0.0 ;  (* graph basis: NUT_TO_BED normal 0.00 L/h )
  FB_PI_NUTRIENT_DOSEFT-02( PV := NUTRIENT_DOSEFT-02_PV, SP := NUTRIENT_DOSEFT-02_SP );  (* PI per AQS-CTL-002; GAIN/KI entered at commissioning from the step test (AQS-COM-001 sec. 3), anti-windup clamp per this FB *)
  NUTRIENT_DOSEFT-02_ALARM_HI := 0.0 ;  (* expected-zero state: any positive PV alarms )

  (* FLOW control loop - set-point from the graph basis *)
  NUTRIENT_DOSEFT-03_SP := 0.58 ;  (* graph basis: IA-NUT-01 normal 0.58 L/h )
  FB_PI_NUTRIENT_DOSEFT-03( PV := NUTRIENT_DOSEFT-03_PV, SP := NUTRIENT_DOSEFT-03_SP );  (* PI per AQS-CTL-002; GAIN/KI entered at commissioning from the step test (AQS-COM-001 sec. 3), anti-windup clamp per this FB *)
  NUTRIENT_DOSEFT-03_ALARM_HI := 0.638 ;  (* SP x 1.1 margin, A-M-188 margin class *)
  NUTRIENT_DOSEFT-03_ALARM_LO := 0.522 ;

  (* FLOW control loop - set-point from the graph basis *)
  NUTRIENT_DOSEFT-04_SP := 3.43 ;  (* graph basis: IA-NUT-LEACH normal 3.43 L/h )
  FB_PI_NUTRIENT_DOSEFT-04( PV := NUTRIENT_DOSEFT-04_PV, SP := NUTRIENT_DOSEFT-04_SP );  (* PI per AQS-CTL-002; GAIN/KI entered at commissioning from the step test (AQS-COM-001 sec. 3), anti-windup clamp per this FB *)
  NUTRIENT_DOSEFT-04_ALARM_HI := 3.7730000000000006 ;  (* SP x 1.1 margin, A-M-188 margin class *)
  NUTRIENT_DOSEFT-04_ALARM_LO := 3.087 ;

  (* FLOW control loop - set-point from the graph basis *)
  NUTRIENT_DOSEFT-05_SP := 1.31 ;  (* graph basis: IA-NUT-BED normal 1.31 L/h )
  FB_PI_NUTRIENT_DOSEFT-05( PV := NUTRIENT_DOSEFT-05_PV, SP := NUTRIENT_DOSEFT-05_SP );  (* PI per AQS-CTL-002; GAIN/KI entered at commissioning from the step test (AQS-COM-001 sec. 3), anti-windup clamp per this FB *)
  NUTRIENT_DOSEFT-05_ALARM_HI := 1.4410000000000003 ;  (* SP x 1.1 margin, A-M-188 margin class *)
  NUTRIENT_DOSEFT-05_ALARM_LO := 1.179 ;

  (* FLOW control loop - set-point from the graph basis *)
  NUTRIENT_DOSEFT-06_SP := 0.02 ;  (* graph basis: IA-SIC-RET normal 0.02 L/h )
  FB_PI_NUTRIENT_DOSEFT-06( PV := NUTRIENT_DOSEFT-06_PV, SP := NUTRIENT_DOSEFT-06_SP );  (* PI per AQS-CTL-002; GAIN/KI entered at commissioning from the step test (AQS-COM-001 sec. 3), anti-windup clamp per this FB *)
  NUTRIENT_DOSEFT-06_ALARM_HI := 0.022000000000000002 ;  (* SP x 1.1 margin, A-M-188 margin class *)
  NUTRIENT_DOSEFT-06_ALARM_LO := 0.018000000000000002 ;

  (* LEVEL monitoring block - indication, no set-point invented )
  FB_AI_NUTRIENT_DOSELT-01( PV := NUTRIENT_DOSELT-01_PV );
  NUTRIENT_DOSELT-01_ALARM_HI := 90.0 ;  (* 90 % of span, registered LSH convention )

  (* PRESSURE monitoring block - indication, no set-point invented )
  FB_AI_NUTRIENT_DOSEPT-01( PV := NUTRIENT_DOSEPT-01_PV );
  NUTRIENT_DOSEPT-01_ALARM_HI := 9.0 ;  (* 90 % of span, registered LSH convention )

  (* TEMPERATURE monitoring block - indication, no set-point invented )
  FB_AI_NUTRIENT_DOSETE-01( PV := NUTRIENT_DOSETE-01_PV );
  NUTRIENT_DOSETE-01_ALARM_HI := 135.0 ;  (* 90 % of span, registered LSH convention )

END_PROGRAM

(* ---- PLC-OIL.st ---- *)
(* AQS-CTL-004 X-CTL-04: control program source, generated by flow_graph/control/plc_programs.py *)
(* Basis: AQS-CTL-001 INSTRUMENT_INDEX.csv, AQS-CTL-002 control architecture, graph set-points. *)
(* PLC-OIL: CPU single; IO counts AI 55 AO 0 DI 33 DO 4 (modules per AQS-CTL-002, 16-channel, 20 % spare) *)
PROGRAM PLC_OIL_CTRL
VAR
  (* 100 ms cyclic task per AQS-CTL-002 *)
  HOPPERFT-01_PV : REAL ;  (* IA-FEED-01 normal 4.28 L/h )
  HOPPERPT-01_PV : REAL ;  (* no design pressure on the graph )
  HOPPERTE-01_PV : REAL ;  (* band by service )
  AFTERBURNERPT-01_PV : REAL ;  (* no design pressure on the graph )
  AFTERBURNERTE-01_PV : REAL ;  (* band by service )
  OIL_DRYERLT-01_PV : REAL ;  (* A-M-182 liquid height )
  OIL_DRYERPT-01_PV : REAL ;  (* no design pressure on the graph )
  OIL_DRYERTE-01_PV : REAL ;  (* band by service )
  OIL_FRACFT-01_PV : REAL ;  (* CUT-1 normal 0.33 L/h )
  OIL_FRACFT-02_PV : REAL ;  (* CUT-2 normal 0.41 L/h )
  OIL_FRACFT-03_PV : REAL ;  (* CUT-3 normal 0.26 L/h )
  OIL_FRACFT-04_PV : REAL ;  (* CUT-4 normal 0.24 L/h )
  OIL_FRACFT-05_PV : REAL ;  (* IA-OIL-03 normal 0.21 L/h )
  OIL_FRACFT-06_PV : REAL ;  (* OIL_TO_OLEFIN normal 0.00 L/h )
  OIL_FRACLT-01_PV : REAL ;  (* A-M-182 liquid height )
  OIL_FRACPT-01_PV : REAL ;  (* no design pressure on the graph )
  OIL_FRACTE-01_PV : REAL ;  (* band by service )
  OIL_PYROFT-01_PV : REAL ;  (* IA-OIL-02 normal 1.39 L/h )
  OIL_PYROLT-01_PV : REAL ;  (* A-M-182 liquid height )
  OIL_PYROPT-01_PV : REAL ;  (* no design pressure on the graph )
  OIL_PYROTE-01_PV : REAL ;  (* design T 500.0 C )
  PROD_C11_C18LT-01_PV : REAL ;  (* A-M-182 liquid height )
  PROD_C11_C18PT-01_PV : REAL ;  (* no design pressure on the graph )
  PROD_C11_C18TE-01_PV : REAL ;  (* band by service )
  PROD_C19_C28FT-01_PV : REAL ;  (* WAX_TO_GREASE_CA normal 0.00 L/h )
  PROD_C19_C28FT-02_PV : REAL ;  (* WAX_TO_GREASE_LI normal 0.00 L/h )
  PROD_C19_C28FT-03_PV : REAL ;  (* CUT-3-OUT normal 0.16 L/h )
  PROD_C19_C28FT-04_PV : REAL ;  (* IA-C19-SHIP normal 0.09 L/h )
  PROD_C19_C28LT-01_PV : REAL ;  (* A-M-182 liquid height )
  PROD_C19_C28PT-01_PV : REAL ;  (* no design pressure on the graph )
  PROD_C19_C28TE-01_PV : REAL ;  (* band by service )
  PROD_C29FT-01_PV : REAL ;  (* C29_RECYCLE normal 0.24 L/h )
  PROD_C29LT-01_PV : REAL ;  (* A-M-182 liquid height )
  PROD_C29PT-01_PV : REAL ;  (* no design pressure on the graph )
  PROD_C29TE-01_PV : REAL ;  (* band by service )
  PROD_C5_C10FT-01_PV : REAL ;  (* CUT-1-OUT normal 0.00 L/h )
  PROD_C5_C10FT-02_PV : REAL ;  (* IA-C5-SHIP normal 0.32 L/h )
  PROD_C5_C10FT-03_PV : REAL ;  (* IA-C5-POLY normal 0.01 L/h )
  PROD_C5_C10LT-01_PV : REAL ;  (* A-M-182 liquid height )
  PROD_C5_C10PT-01_PV : REAL ;  (* no design pressure on the graph )
  PROD_C5_C10TE-01_PV : REAL ;  (* band by service )
  GREASE_CALT-01_PV : REAL ;  (* A-M-182 liquid height )
  GREASE_CAPT-01_PV : REAL ;  (* no design pressure on the graph )
  GREASE_CATE-01_PV : REAL ;  (* band by service )
  GREASE_LIPT-01_PV : REAL ;  (* no design pressure on the graph )
  GREASE_LITE-01_PV : REAL ;  (* band by service )
  C29_RECYCLELT-01_PV : REAL ;  (* A-M-182 liquid height )
  C29_RECYCLEPT-01_PV : REAL ;  (* no design pressure on the graph )
  C29_RECYCLETE-01_PV : REAL ;  (* band by service )
  NCG_HEADERPT-01_PV : REAL ;  (* NCG header: IA-OIL-03 5.0 kg/d to the afterburner; no design pressure on the gra )
  GREASE_LILT-01_PV : REAL ;  (* kettle holdup (class kettle) )
  CAT_OXTE-01_PV : REAL ;  (* catalyst bed temperature watch against the A-M-399 450 C light-off window (X-LOC )
  AFTERBURNERTE-90 : BOOL ;  (* SIF watch input, routed to the safety CPU pair (AQS-CTL-003) *)
  OIL_DRYERTE-90 : BOOL ;  (* SIF watch input, routed to the safety CPU pair (AQS-CTL-003) *)
  OIL_PYROTE-90 : BOOL ;  (* SIF watch input, routed to the safety CPU pair (AQS-CTL-003) *)
END_VAR

  (* FLOW control loop - set-point from the graph basis *)
  HOPPERFT-01_SP := 4.28 ;  (* graph basis: IA-FEED-01 normal 4.28 L/h )
  FB_PI_HOPPERFT-01( PV := HOPPERFT-01_PV, SP := HOPPERFT-01_SP );  (* PI per AQS-CTL-002; GAIN/KI entered at commissioning from the step test (AQS-COM-001 sec. 3), anti-windup clamp per this FB *)
  HOPPERFT-01_ALARM_HI := 4.708000000000001 ;  (* SP x 1.1 margin, A-M-188 margin class *)
  HOPPERFT-01_ALARM_LO := 3.8520000000000003 ;

  (* PRESSURE monitoring block - indication, no set-point invented )
  FB_AI_HOPPERPT-01( PV := HOPPERPT-01_PV );
  HOPPERPT-01_ALARM_HI := 9.0 ;  (* 90 % of span, registered LSH convention )

  (* TEMPERATURE monitoring block - indication, no set-point invented )
  FB_AI_HOPPERTE-01( PV := HOPPERTE-01_PV );
  HOPPERTE-01_ALARM_HI := 135.0 ;  (* 90 % of span, registered LSH convention )

  (* PRESSURE monitoring block - indication, no set-point invented )
  FB_AI_AFTERBURNERPT-01( PV := AFTERBURNERPT-01_PV );
  AFTERBURNERPT-01_ALARM_HI := 9.0 ;  (* 90 % of span, registered LSH convention )

  (* TEMPERATURE monitoring block - indication, no set-point invented )
  FB_AI_AFTERBURNERTE-01( PV := AFTERBURNERTE-01_PV );
  AFTERBURNERTE-01_ALARM_HI := 540.0 ;  (* 90 % of span, registered LSH convention )

  (* LEVEL monitoring block - indication, no set-point invented )
  FB_AI_OIL_DRYERLT-01( PV := OIL_DRYERLT-01_PV );
  OIL_DRYERLT-01_ALARM_HI := 90.0 ;  (* 90 % of span, registered LSH convention )

  (* PRESSURE monitoring block - indication, no set-point invented )
  FB_AI_OIL_DRYERPT-01( PV := OIL_DRYERPT-01_PV );
  OIL_DRYERPT-01_ALARM_HI := 9.0 ;  (* 90 % of span, registered LSH convention )

  (* TEMPERATURE monitoring block - indication, no set-point invented )
  FB_AI_OIL_DRYERTE-01( PV := OIL_DRYERTE-01_PV );
  OIL_DRYERTE-01_ALARM_HI := 540.0 ;  (* 90 % of span, registered LSH convention )

  (* FLOW control loop - set-point from the graph basis *)
  OIL_FRACFT-01_SP := 0.33 ;  (* graph basis: CUT-1 normal 0.33 L/h )
  FB_PI_OIL_FRACFT-01( PV := OIL_FRACFT-01_PV, SP := OIL_FRACFT-01_SP );  (* PI per AQS-CTL-002; GAIN/KI entered at commissioning from the step test (AQS-COM-001 sec. 3), anti-windup clamp per this FB *)
  OIL_FRACFT-01_ALARM_HI := 0.36300000000000004 ;  (* SP x 1.1 margin, A-M-188 margin class *)
  OIL_FRACFT-01_ALARM_LO := 0.29700000000000004 ;

  (* FLOW control loop - set-point from the graph basis *)
  OIL_FRACFT-02_SP := 0.41 ;  (* graph basis: CUT-2 normal 0.41 L/h )
  FB_PI_OIL_FRACFT-02( PV := OIL_FRACFT-02_PV, SP := OIL_FRACFT-02_SP );  (* PI per AQS-CTL-002; GAIN/KI entered at commissioning from the step test (AQS-COM-001 sec. 3), anti-windup clamp per this FB *)
  OIL_FRACFT-02_ALARM_HI := 0.451 ;  (* SP x 1.1 margin, A-M-188 margin class *)
  OIL_FRACFT-02_ALARM_LO := 0.369 ;

  (* FLOW control loop - set-point from the graph basis *)
  OIL_FRACFT-03_SP := 0.26 ;  (* graph basis: CUT-3 normal 0.26 L/h )
  FB_PI_OIL_FRACFT-03( PV := OIL_FRACFT-03_PV, SP := OIL_FRACFT-03_SP );  (* PI per AQS-CTL-002; GAIN/KI entered at commissioning from the step test (AQS-COM-001 sec. 3), anti-windup clamp per this FB *)
  OIL_FRACFT-03_ALARM_HI := 0.28600000000000003 ;  (* SP x 1.1 margin, A-M-188 margin class *)
  OIL_FRACFT-03_ALARM_LO := 0.234 ;

  (* FLOW control loop - set-point from the graph basis *)
  OIL_FRACFT-04_SP := 0.24 ;  (* graph basis: CUT-4 normal 0.24 L/h )
  FB_PI_OIL_FRACFT-04( PV := OIL_FRACFT-04_PV, SP := OIL_FRACFT-04_SP );  (* PI per AQS-CTL-002; GAIN/KI entered at commissioning from the step test (AQS-COM-001 sec. 3), anti-windup clamp per this FB *)
  OIL_FRACFT-04_ALARM_HI := 0.264 ;  (* SP x 1.1 margin, A-M-188 margin class *)
  OIL_FRACFT-04_ALARM_LO := 0.216 ;

  (* FLOW control loop - set-point from the graph basis *)
  OIL_FRACFT-05_SP := 0.21 ;  (* graph basis: IA-OIL-03 normal 0.21 L/h )
  FB_PI_OIL_FRACFT-05( PV := OIL_FRACFT-05_PV, SP := OIL_FRACFT-05_SP );  (* PI per AQS-CTL-002; GAIN/KI entered at commissioning from the step test (AQS-COM-001 sec. 3), anti-windup clamp per this FB *)
  OIL_FRACFT-05_ALARM_HI := 0.231 ;  (* SP x 1.1 margin, A-M-188 margin class *)
  OIL_FRACFT-05_ALARM_LO := 0.189 ;

  (* FLOW control loop - set-point from the graph basis *)
  OIL_FRACFT-06_SP := 0.0 ;  (* graph basis: OIL_TO_OLEFIN normal 0.00 L/h )
  FB_PI_OIL_FRACFT-06( PV := OIL_FRACFT-06_PV, SP := OIL_FRACFT-06_SP );  (* PI per AQS-CTL-002; GAIN/KI entered at commissioning from the step test (AQS-COM-001 sec. 3), anti-windup clamp per this FB *)
  OIL_FRACFT-06_ALARM_HI := 0.0 ;  (* expected-zero state: any positive PV alarms )

  (* LEVEL monitoring block - indication, no set-point invented )
  FB_AI_OIL_FRACLT-01( PV := OIL_FRACLT-01_PV );
  OIL_FRACLT-01_ALARM_HI := 90.0 ;  (* 90 % of span, registered LSH convention )

  (* PRESSURE monitoring block - indication, no set-point invented )
  FB_AI_OIL_FRACPT-01( PV := OIL_FRACPT-01_PV );
  OIL_FRACPT-01_ALARM_HI := 9.0 ;  (* 90 % of span, registered LSH convention )

  (* TEMPERATURE monitoring block - indication, no set-point invented )
  FB_AI_OIL_FRACTE-01( PV := OIL_FRACTE-01_PV );
  OIL_FRACTE-01_ALARM_HI := 135.0 ;  (* 90 % of span, registered LSH convention )

  (* FLOW control loop - set-point from the graph basis *)
  OIL_PYROFT-01_SP := 1.39 ;  (* graph basis: IA-OIL-02 normal 1.39 L/h )
  FB_PI_OIL_PYROFT-01( PV := OIL_PYROFT-01_PV, SP := OIL_PYROFT-01_SP );  (* PI per AQS-CTL-002; GAIN/KI entered at commissioning from the step test (AQS-COM-001 sec. 3), anti-windup clamp per this FB *)
  OIL_PYROFT-01_ALARM_HI := 1.529 ;  (* SP x 1.1 margin, A-M-188 margin class *)
  OIL_PYROFT-01_ALARM_LO := 1.251 ;

  (* LEVEL monitoring block - indication, no set-point invented )
  FB_AI_OIL_PYROLT-01( PV := OIL_PYROLT-01_PV );
  OIL_PYROLT-01_ALARM_HI := 90.0 ;  (* 90 % of span, registered LSH convention )

  (* PRESSURE monitoring block - indication, no set-point invented )
  FB_AI_OIL_PYROPT-01( PV := OIL_PYROPT-01_PV );
  OIL_PYROPT-01_ALARM_HI := 9.0 ;  (* 90 % of span, registered LSH convention )

  (* TEMPERATURE control loop - set-point from the graph basis *)
  OIL_PYROTE-01_SP := 500.0 ;  (* graph basis: design T 500.0 C )
  FB_PI_OIL_PYROTE-01( PV := OIL_PYROTE-01_PV, SP := OIL_PYROTE-01_SP );  (* PI per AQS-CTL-002; GAIN/KI entered at commissioning from the step test (AQS-COM-001 sec. 3), anti-windup clamp per this FB *)
  OIL_PYROTE-01_ALARM_HI := 550.0 ;  (* SP x 1.1 margin, A-M-188 margin class *)
  OIL_PYROTE-01_ALARM_LO := 450.0 ;

  (* LEVEL monitoring block - indication, no set-point invented )
  FB_AI_PROD_C11_C18LT-01( PV := PROD_C11_C18LT-01_PV );
  PROD_C11_C18LT-01_ALARM_HI := 90.0 ;  (* 90 % of span, registered LSH convention )

  (* PRESSURE monitoring block - indication, no set-point invented )
  FB_AI_PROD_C11_C18PT-01( PV := PROD_C11_C18PT-01_PV );
  PROD_C11_C18PT-01_ALARM_HI := 9.0 ;  (* 90 % of span, registered LSH convention )

  (* TEMPERATURE monitoring block - indication, no set-point invented )
  FB_AI_PROD_C11_C18TE-01( PV := PROD_C11_C18TE-01_PV );
  PROD_C11_C18TE-01_ALARM_HI := 135.0 ;  (* 90 % of span, registered LSH convention )

  (* FLOW control loop - set-point from the graph basis *)
  PROD_C19_C28FT-01_SP := 0.0 ;  (* graph basis: WAX_TO_GREASE_CA normal 0.00 L/h )
  FB_PI_PROD_C19_C28FT-01( PV := PROD_C19_C28FT-01_PV, SP := PROD_C19_C28FT-01_SP );  (* PI per AQS-CTL-002; GAIN/KI entered at commissioning from the step test (AQS-COM-001 sec. 3), anti-windup clamp per this FB *)
  PROD_C19_C28FT-01_ALARM_HI := 0.0 ;  (* expected-zero state: any positive PV alarms )

  (* FLOW control loop - set-point from the graph basis *)
  PROD_C19_C28FT-02_SP := 0.0 ;  (* graph basis: WAX_TO_GREASE_LI normal 0.00 L/h )
  FB_PI_PROD_C19_C28FT-02( PV := PROD_C19_C28FT-02_PV, SP := PROD_C19_C28FT-02_SP );  (* PI per AQS-CTL-002; GAIN/KI entered at commissioning from the step test (AQS-COM-001 sec. 3), anti-windup clamp per this FB *)
  PROD_C19_C28FT-02_ALARM_HI := 0.0 ;  (* expected-zero state: any positive PV alarms )

  (* FLOW control loop - set-point from the graph basis *)
  PROD_C19_C28FT-03_SP := 0.16 ;  (* graph basis: CUT-3-OUT normal 0.16 L/h )
  FB_PI_PROD_C19_C28FT-03( PV := PROD_C19_C28FT-03_PV, SP := PROD_C19_C28FT-03_SP );  (* PI per AQS-CTL-002; GAIN/KI entered at commissioning from the step test (AQS-COM-001 sec. 3), anti-windup clamp per this FB *)
  PROD_C19_C28FT-03_ALARM_HI := 0.17600000000000002 ;  (* SP x 1.1 margin, A-M-188 margin class *)
  PROD_C19_C28FT-03_ALARM_LO := 0.14400000000000002 ;

  (* FLOW control loop - set-point from the graph basis *)
  PROD_C19_C28FT-04_SP := 0.09 ;  (* graph basis: IA-C19-SHIP normal 0.09 L/h )
  FB_PI_PROD_C19_C28FT-04( PV := PROD_C19_C28FT-04_PV, SP := PROD_C19_C28FT-04_SP );  (* PI per AQS-CTL-002; GAIN/KI entered at commissioning from the step test (AQS-COM-001 sec. 3), anti-windup clamp per this FB *)
  PROD_C19_C28FT-04_ALARM_HI := 0.099 ;  (* SP x 1.1 margin, A-M-188 margin class *)
  PROD_C19_C28FT-04_ALARM_LO := 0.081 ;

  (* LEVEL monitoring block - indication, no set-point invented )
  FB_AI_PROD_C19_C28LT-01( PV := PROD_C19_C28LT-01_PV );
  PROD_C19_C28LT-01_ALARM_HI := 90.0 ;  (* 90 % of span, registered LSH convention )

  (* PRESSURE monitoring block - indication, no set-point invented )
  FB_AI_PROD_C19_C28PT-01( PV := PROD_C19_C28PT-01_PV );
  PROD_C19_C28PT-01_ALARM_HI := 9.0 ;  (* 90 % of span, registered LSH convention )

  (* TEMPERATURE monitoring block - indication, no set-point invented )
  FB_AI_PROD_C19_C28TE-01( PV := PROD_C19_C28TE-01_PV );
  PROD_C19_C28TE-01_ALARM_HI := 135.0 ;  (* 90 % of span, registered LSH convention )

  (* FLOW control loop - set-point from the graph basis *)
  PROD_C29FT-01_SP := 0.24 ;  (* graph basis: C29_RECYCLE normal 0.24 L/h )
  FB_PI_PROD_C29FT-01( PV := PROD_C29FT-01_PV, SP := PROD_C29FT-01_SP );  (* PI per AQS-CTL-002; GAIN/KI entered at commissioning from the step test (AQS-COM-001 sec. 3), anti-windup clamp per this FB *)
  PROD_C29FT-01_ALARM_HI := 0.264 ;  (* SP x 1.1 margin, A-M-188 margin class *)
  PROD_C29FT-01_ALARM_LO := 0.216 ;

  (* LEVEL monitoring block - indication, no set-point invented )
  FB_AI_PROD_C29LT-01( PV := PROD_C29LT-01_PV );
  PROD_C29LT-01_ALARM_HI := 90.0 ;  (* 90 % of span, registered LSH convention )

  (* PRESSURE monitoring block - indication, no set-point invented )
  FB_AI_PROD_C29PT-01( PV := PROD_C29PT-01_PV );
  PROD_C29PT-01_ALARM_HI := 9.0 ;  (* 90 % of span, registered LSH convention )

  (* TEMPERATURE monitoring block - indication, no set-point invented )
  FB_AI_PROD_C29TE-01( PV := PROD_C29TE-01_PV );
  PROD_C29TE-01_ALARM_HI := 135.0 ;  (* 90 % of span, registered LSH convention )

  (* FLOW control loop - set-point from the graph basis *)
  PROD_C5_C10FT-01_SP := 0.0 ;  (* graph basis: CUT-1-OUT normal 0.00 L/h )
  FB_PI_PROD_C5_C10FT-01( PV := PROD_C5_C10FT-01_PV, SP := PROD_C5_C10FT-01_SP );  (* PI per AQS-CTL-002; GAIN/KI entered at commissioning from the step test (AQS-COM-001 sec. 3), anti-windup clamp per this FB *)
  PROD_C5_C10FT-01_ALARM_HI := 0.0 ;  (* expected-zero state: any positive PV alarms )

  (* FLOW control loop - set-point from the graph basis *)
  PROD_C5_C10FT-02_SP := 0.32 ;  (* graph basis: IA-C5-SHIP normal 0.32 L/h )
  FB_PI_PROD_C5_C10FT-02( PV := PROD_C5_C10FT-02_PV, SP := PROD_C5_C10FT-02_SP );  (* PI per AQS-CTL-002; GAIN/KI entered at commissioning from the step test (AQS-COM-001 sec. 3), anti-windup clamp per this FB *)
  PROD_C5_C10FT-02_ALARM_HI := 0.35200000000000004 ;  (* SP x 1.1 margin, A-M-188 margin class *)
  PROD_C5_C10FT-02_ALARM_LO := 0.28800000000000003 ;

  (* FLOW control loop - set-point from the graph basis *)
  PROD_C5_C10FT-03_SP := 0.01 ;  (* graph basis: IA-C5-POLY normal 0.01 L/h )
  FB_PI_PROD_C5_C10FT-03( PV := PROD_C5_C10FT-03_PV, SP := PROD_C5_C10FT-03_SP );  (* PI per AQS-CTL-002; GAIN/KI entered at commissioning from the step test (AQS-COM-001 sec. 3), anti-windup clamp per this FB *)
  PROD_C5_C10FT-03_ALARM_HI := 0.011000000000000001 ;  (* SP x 1.1 margin, A-M-188 margin class *)
  PROD_C5_C10FT-03_ALARM_LO := 0.009000000000000001 ;

  (* LEVEL monitoring block - indication, no set-point invented )
  FB_AI_PROD_C5_C10LT-01( PV := PROD_C5_C10LT-01_PV );
  PROD_C5_C10LT-01_ALARM_HI := 90.0 ;  (* 90 % of span, registered LSH convention )

  (* PRESSURE monitoring block - indication, no set-point invented )
  FB_AI_PROD_C5_C10PT-01( PV := PROD_C5_C10PT-01_PV );
  PROD_C5_C10PT-01_ALARM_HI := 9.0 ;  (* 90 % of span, registered LSH convention )

  (* TEMPERATURE monitoring block - indication, no set-point invented )
  FB_AI_PROD_C5_C10TE-01( PV := PROD_C5_C10TE-01_PV );
  PROD_C5_C10TE-01_ALARM_HI := 135.0 ;  (* 90 % of span, registered LSH convention )

  (* LEVEL monitoring block - indication, no set-point invented )
  FB_AI_GREASE_CALT-01( PV := GREASE_CALT-01_PV );
  GREASE_CALT-01_ALARM_HI := 90.0 ;  (* 90 % of span, registered LSH convention )

  (* PRESSURE monitoring block - indication, no set-point invented )
  FB_AI_GREASE_CAPT-01( PV := GREASE_CAPT-01_PV );
  GREASE_CAPT-01_ALARM_HI := 9.0 ;  (* 90 % of span, registered LSH convention )

  (* TEMPERATURE monitoring block - indication, no set-point invented )
  FB_AI_GREASE_CATE-01( PV := GREASE_CATE-01_PV );
  GREASE_CATE-01_ALARM_HI := 135.0 ;  (* 90 % of span, registered LSH convention )

  (* PRESSURE monitoring block - indication, no set-point invented )
  FB_AI_GREASE_LIPT-01( PV := GREASE_LIPT-01_PV );
  GREASE_LIPT-01_ALARM_HI := 9.0 ;  (* 90 % of span, registered LSH convention )

  (* TEMPERATURE monitoring block - indication, no set-point invented )
  FB_AI_GREASE_LITE-01( PV := GREASE_LITE-01_PV );
  GREASE_LITE-01_ALARM_HI := 135.0 ;  (* 90 % of span, registered LSH convention )

  (* LEVEL monitoring block - indication, no set-point invented )
  FB_AI_C29_RECYCLELT-01( PV := C29_RECYCLELT-01_PV );
  C29_RECYCLELT-01_ALARM_HI := 90.0 ;  (* 90 % of span, registered LSH convention )

  (* PRESSURE monitoring block - indication, no set-point invented )
  FB_AI_C29_RECYCLEPT-01( PV := C29_RECYCLEPT-01_PV );
  C29_RECYCLEPT-01_ALARM_HI := 9.0 ;  (* 90 % of span, registered LSH convention )

  (* TEMPERATURE monitoring block - indication, no set-point invented )
  FB_AI_C29_RECYCLETE-01( PV := C29_RECYCLETE-01_PV );
  C29_RECYCLETE-01_ALARM_HI := 135.0 ;  (* 90 % of span, registered LSH convention )

  (* PRESSURE monitoring block - indication, no set-point invented )
  FB_AI_NCG_HEADERPT-01( PV := NCG_HEADERPT-01_PV );
  NCG_HEADERPT-01_ALARM_HI := 9.0 ;  (* 90 % of span, registered LSH convention )

  (* LEVEL monitoring block - indication, no set-point invented )
  FB_AI_GREASE_LILT-01( PV := GREASE_LILT-01_PV );
  GREASE_LILT-01_ALARM_HI := 90.0 ;  (* 90 % of span, registered LSH convention )

  (* TEMPERATURE monitoring block - indication, no set-point invented )
  FB_AI_CAT_OXTE-01( PV := CAT_OXTE-01_PV );
  CAT_OXTE-01_ALARM_HI := 540.0 ;  (* 90 % of span, registered LSH convention )

  (* SIF watch passthrough, no action in the basic program )
  SIF_WATCH_AFTERBURNERTE-90 := AFTERBURNERTE-90 ;  (* to safety CPU pair, AQS-CTL-003 )

  (* SIF watch passthrough, no action in the basic program )
  SIF_WATCH_OIL_DRYERTE-90 := OIL_DRYERTE-90 ;  (* to safety CPU pair, AQS-CTL-003 )

  (* SIF watch passthrough, no action in the basic program )
  SIF_WATCH_OIL_PYROTE-90 := OIL_PYROTE-90 ;  (* to safety CPU pair, AQS-CTL-003 )

END_PROGRAM

(* ---- PLC-POLYMERS.st ---- *)
(* AQS-CTL-004 X-CTL-04: control program source, generated by flow_graph/control/plc_programs.py *)
(* Basis: AQS-CTL-001 INSTRUMENT_INDEX.csv, AQS-CTL-002 control architecture, graph set-points. *)
(* PLC-POLYMERS: CPU single; IO counts AI 53 AO 0 DI 27 DO 5 (modules per AQS-CTL-002, 16-channel, 20 % spare) *)
PROGRAM PLC_POLYMERS_CTRL
VAR
  (* 100 ms cyclic task per AQS-CTL-002 *)
  FILM_CASTLT-01_PV : REAL ;  (* A-M-182 liquid height )
  FILM_CASTPT-01_PV : REAL ;  (* no design pressure on the graph )
  FILM_CASTTE-01_PV : REAL ;  (* band by service )
  HF_GENFT-01_PV : REAL ;  (* HF_GEN_TO_VDF normal 0.00 L/h )
  HF_GENFT-02_PV : REAL ;  (* HF_GEN_TO_TFE normal 0.00 L/h )
  HF_GENFT-03_PV : REAL ;  (* IA-HF-PROD normal 0.06 L/h )
  HF_GENLT-01_PV : REAL ;  (* A-M-182 liquid height )
  HF_GENPT-01_PV : REAL ;  (* no design pressure on the graph )
  HF_GENTE-01_PV : REAL ;  (* design T 250.0 C )
  PELLETPT-01_PV : REAL ;  (* no design pressure on the graph )
  PELLETTE-01_PV : REAL ;  (* band by service )
  POLY_CONDPT-01_PV : REAL ;  (* no design pressure on the graph )
  POLY_CONDTE-01_PV : REAL ;  (* band by service )
  POLY_FFT-01_PV : REAL ;  (* POLYF_TO_FILM normal 0.01 L/h )
  POLY_FFT-02_PV : REAL ;  (* POLYF_RECLAIM normal 0.00 L/h )
  POLY_FLT-01_PV : REAL ;  (* A-M-182 liquid height )
  POLY_FPT-01_PV : REAL ;  (* no design pressure on the graph )
  POLY_FTE-01_PV : REAL ;  (* design T 60 C )
  POLY_OLEFINLT-01_PV : REAL ;  (* A-M-182 liquid height )
  POLY_OLEFINPT-01_PV : REAL ;  (* design 5000.0 kPa g )
  POLY_OLEFINTE-01_PV : REAL ;  (* design T 250.0 C )
  POLY_STOCKFT-01_PV : REAL ;  (* FLUORO_TO_MFG normal 0.01 L/h )
  POLY_STOCKFT-02_PV : REAL ;  (* STOCK_TO_FIBER normal 0.00 L/h )
  POLY_STOCKPT-01_PV : REAL ;  (* no design pressure on the graph )
  POLY_STOCKTE-01_PV : REAL ;  (* band by service )
  POWDER_RESINPT-01_PV : REAL ;  (* no design pressure on the graph )
  POWDER_RESINTE-01_PV : REAL ;  (* band by service )
  TFE_SYNFT-01_PV : REAL ;  (* TFE_TO_POLY_F normal 0.00 L/h )
  TFE_SYNFT-02_PV : REAL ;  (* TFE_HCL_TO_CRU normal 0.01 L/h )
  TFE_SYNLT-01_PV : REAL ;  (* A-M-182 liquid height )
  TFE_SYNPT-01_PV : REAL ;  (* no design pressure on the graph )
  TFE_SYNTE-01_PV : REAL ;  (* band by service )
  VDF_SYNFT-01_PV : REAL ;  (* VDF_TO_POLY_F normal 0.01 L/h )
  VDF_SYNFT-02_PV : REAL ;  (* VDF_HCL_TO_CRU normal 0.02 L/h )
  VDF_SYNLT-01_PV : REAL ;  (* A-M-182 liquid height )
  VDF_SYNPT-01_PV : REAL ;  (* no design pressure on the graph )
  VDF_SYNTE-01_PV : REAL ;  (* band by service )
  POLY_FIBERFT-01_PV : REAL ;  (* FIBER_SCRAP normal 0.00 L/h )
  POLY_FIBERFT-02_PV : REAL ;  (* FLEECE_TO_MFG normal 0.00 L/h )
  POLY_FIBERPT-01_PV : REAL ;  (* no design pressure on the graph )
  POLY_FIBERTE-01_PV : REAL ;  (* band by service )
  ACID_PLANTLT-01_PV : REAL ;  (* A-M-182 liquid height )
  ACID_PLANTPT-01_PV : REAL ;  (* no design pressure on the graph )
  ACID_PLANTTE-01_PV : REAL ;  (* band by service )
  HF_GENAE-01_PV : REAL ;  (* kiln offgas HF watch: design hf_kg_d 1.67 kg/d )
  POLY_CONDLT-01_PV : REAL ;  (* kettle: design H_mm 300 )
  POWDER_RESINST-01_PV : REAL ;  (* mill drive: design duty_kW 0.0152 kW )
  FILM_CASTST-01_PV : REAL ;  (* chill-roll drive: design chill_roll_D_mm 150 )
  POLY_STOCKLT-01_PV : REAL ;  (* pellet tote bins (design bin) )
  POLY_FIBERTIR-01_PV : REAL ;  (* melt temperature is the spin-quality variable: PP spins at the 200-260 C class ( )
  POLY_FIBERFIT-01_PV : REAL ;  (* denier control: fibre mass per unit length follows the pump volumetric consisten )
  HF_GENTE-90 : BOOL ;  (* SIF watch input, routed to the safety CPU pair (AQS-CTL-003) *)
  POLY_OLEFINTE-90 : BOOL ;  (* SIF watch input, routed to the safety CPU pair (AQS-CTL-003) *)
END_VAR

  (* LEVEL monitoring block - indication, no set-point invented )
  FB_AI_FILM_CASTLT-01( PV := FILM_CASTLT-01_PV );
  FILM_CASTLT-01_ALARM_HI := 90.0 ;  (* 90 % of span, registered LSH convention )

  (* PRESSURE monitoring block - indication, no set-point invented )
  FB_AI_FILM_CASTPT-01( PV := FILM_CASTPT-01_PV );
  FILM_CASTPT-01_ALARM_HI := 9.0 ;  (* 90 % of span, registered LSH convention )

  (* TEMPERATURE monitoring block - indication, no set-point invented )
  FB_AI_FILM_CASTTE-01( PV := FILM_CASTTE-01_PV );
  FILM_CASTTE-01_ALARM_HI := 135.0 ;  (* 90 % of span, registered LSH convention )

  (* FLOW control loop - set-point from the graph basis *)
  HF_GENFT-01_SP := 0.0 ;  (* graph basis: HF_GEN_TO_VDF normal 0.00 L/h )
  FB_PI_HF_GENFT-01( PV := HF_GENFT-01_PV, SP := HF_GENFT-01_SP );  (* PI per AQS-CTL-002; GAIN/KI entered at commissioning from the step test (AQS-COM-001 sec. 3), anti-windup clamp per this FB *)
  HF_GENFT-01_ALARM_HI := 0.0 ;  (* expected-zero state: any positive PV alarms )

  (* FLOW control loop - set-point from the graph basis *)
  HF_GENFT-02_SP := 0.0 ;  (* graph basis: HF_GEN_TO_TFE normal 0.00 L/h )
  FB_PI_HF_GENFT-02( PV := HF_GENFT-02_PV, SP := HF_GENFT-02_SP );  (* PI per AQS-CTL-002; GAIN/KI entered at commissioning from the step test (AQS-COM-001 sec. 3), anti-windup clamp per this FB *)
  HF_GENFT-02_ALARM_HI := 0.0 ;  (* expected-zero state: any positive PV alarms )

  (* FLOW control loop - set-point from the graph basis *)
  HF_GENFT-03_SP := 0.06 ;  (* graph basis: IA-HF-PROD normal 0.06 L/h )
  FB_PI_HF_GENFT-03( PV := HF_GENFT-03_PV, SP := HF_GENFT-03_SP );  (* PI per AQS-CTL-002; GAIN/KI entered at commissioning from the step test (AQS-COM-001 sec. 3), anti-windup clamp per this FB *)
  HF_GENFT-03_ALARM_HI := 0.066 ;  (* SP x 1.1 margin, A-M-188 margin class *)
  HF_GENFT-03_ALARM_LO := 0.054 ;

  (* LEVEL monitoring block - indication, no set-point invented )
  FB_AI_HF_GENLT-01( PV := HF_GENLT-01_PV );
  HF_GENLT-01_ALARM_HI := 90.0 ;  (* 90 % of span, registered LSH convention )

  (* PRESSURE monitoring block - indication, no set-point invented )
  FB_AI_HF_GENPT-01( PV := HF_GENPT-01_PV );
  HF_GENPT-01_ALARM_HI := 9.0 ;  (* 90 % of span, registered LSH convention )

  (* TEMPERATURE control loop - set-point from the graph basis *)
  HF_GENTE-01_SP := 250.0 ;  (* graph basis: design T 250.0 C )
  FB_PI_HF_GENTE-01( PV := HF_GENTE-01_PV, SP := HF_GENTE-01_SP );  (* PI per AQS-CTL-002; GAIN/KI entered at commissioning from the step test (AQS-COM-001 sec. 3), anti-windup clamp per this FB *)
  HF_GENTE-01_ALARM_HI := 275.0 ;  (* SP x 1.1 margin, A-M-188 margin class *)
  HF_GENTE-01_ALARM_LO := 225.0 ;

  (* PRESSURE monitoring block - indication, no set-point invented )
  FB_AI_PELLETPT-01( PV := PELLETPT-01_PV );
  PELLETPT-01_ALARM_HI := 9.0 ;  (* 90 % of span, registered LSH convention )

  (* TEMPERATURE monitoring block - indication, no set-point invented )
  FB_AI_PELLETTE-01( PV := PELLETTE-01_PV );
  PELLETTE-01_ALARM_HI := 135.0 ;  (* 90 % of span, registered LSH convention )

  (* PRESSURE monitoring block - indication, no set-point invented )
  FB_AI_POLY_CONDPT-01( PV := POLY_CONDPT-01_PV );
  POLY_CONDPT-01_ALARM_HI := 9.0 ;  (* 90 % of span, registered LSH convention )

  (* TEMPERATURE monitoring block - indication, no set-point invented )
  FB_AI_POLY_CONDTE-01( PV := POLY_CONDTE-01_PV );
  POLY_CONDTE-01_ALARM_HI := 135.0 ;  (* 90 % of span, registered LSH convention )

  (* FLOW control loop - set-point from the graph basis *)
  POLY_FFT-01_SP := 0.01 ;  (* graph basis: POLYF_TO_FILM normal 0.01 L/h )
  FB_PI_POLY_FFT-01( PV := POLY_FFT-01_PV, SP := POLY_FFT-01_SP );  (* PI per AQS-CTL-002; GAIN/KI entered at commissioning from the step test (AQS-COM-001 sec. 3), anti-windup clamp per this FB *)
  POLY_FFT-01_ALARM_HI := 0.011000000000000001 ;  (* SP x 1.1 margin, A-M-188 margin class *)
  POLY_FFT-01_ALARM_LO := 0.009000000000000001 ;

  (* FLOW control loop - set-point from the graph basis *)
  POLY_FFT-02_SP := 0.0 ;  (* graph basis: POLYF_RECLAIM normal 0.00 L/h )
  FB_PI_POLY_FFT-02( PV := POLY_FFT-02_PV, SP := POLY_FFT-02_SP );  (* PI per AQS-CTL-002; GAIN/KI entered at commissioning from the step test (AQS-COM-001 sec. 3), anti-windup clamp per this FB *)
  POLY_FFT-02_ALARM_HI := 0.0 ;  (* expected-zero state: any positive PV alarms )

  (* LEVEL monitoring block - indication, no set-point invented )
  FB_AI_POLY_FLT-01( PV := POLY_FLT-01_PV );
  POLY_FLT-01_ALARM_HI := 90.0 ;  (* 90 % of span, registered LSH convention )

  (* PRESSURE monitoring block - indication, no set-point invented )
  FB_AI_POLY_FPT-01( PV := POLY_FPT-01_PV );
  POLY_FPT-01_ALARM_HI := 9.0 ;  (* 90 % of span, registered LSH convention )

  (* TEMPERATURE control loop - set-point from the graph basis *)
  POLY_FTE-01_SP := 60.0 ;  (* graph basis: design T 60 C )
  FB_PI_POLY_FTE-01( PV := POLY_FTE-01_PV, SP := POLY_FTE-01_SP );  (* PI per AQS-CTL-002; GAIN/KI entered at commissioning from the step test (AQS-COM-001 sec. 3), anti-windup clamp per this FB *)
  POLY_FTE-01_ALARM_HI := 66.0 ;  (* SP x 1.1 margin, A-M-188 margin class *)
  POLY_FTE-01_ALARM_LO := 54.0 ;

  (* LEVEL monitoring block - indication, no set-point invented )
  FB_AI_POLY_OLEFINLT-01( PV := POLY_OLEFINLT-01_PV );
  POLY_OLEFINLT-01_ALARM_HI := 90.0 ;  (* 90 % of span, registered LSH convention )

  (* PRESSURE control loop - set-point from the graph basis *)
  POLY_OLEFINPT-01_SP := 5000.0 ;  (* graph basis: design 5000.0 kPa g )
  FB_PI_POLY_OLEFINPT-01( PV := POLY_OLEFINPT-01_PV, SP := POLY_OLEFINPT-01_SP );  (* PI per AQS-CTL-002; GAIN/KI entered at commissioning from the step test (AQS-COM-001 sec. 3), anti-windup clamp per this FB *)
  POLY_OLEFINPT-01_ALARM_HI := 5500.0 ;  (* SP x 1.1 margin, A-M-188 margin class *)
  POLY_OLEFINPT-01_ALARM_LO := 4500.0 ;

  (* TEMPERATURE control loop - set-point from the graph basis *)
  POLY_OLEFINTE-01_SP := 250.0 ;  (* graph basis: design T 250.0 C )
  FB_PI_POLY_OLEFINTE-01( PV := POLY_OLEFINTE-01_PV, SP := POLY_OLEFINTE-01_SP );  (* PI per AQS-CTL-002; GAIN/KI entered at commissioning from the step test (AQS-COM-001 sec. 3), anti-windup clamp per this FB *)
  POLY_OLEFINTE-01_ALARM_HI := 275.0 ;  (* SP x 1.1 margin, A-M-188 margin class *)
  POLY_OLEFINTE-01_ALARM_LO := 225.0 ;

  (* FLOW control loop - set-point from the graph basis *)
  POLY_STOCKFT-01_SP := 0.01 ;  (* graph basis: FLUORO_TO_MFG normal 0.01 L/h )
  FB_PI_POLY_STOCKFT-01( PV := POLY_STOCKFT-01_PV, SP := POLY_STOCKFT-01_SP );  (* PI per AQS-CTL-002; GAIN/KI entered at commissioning from the step test (AQS-COM-001 sec. 3), anti-windup clamp per this FB *)
  POLY_STOCKFT-01_ALARM_HI := 0.011000000000000001 ;  (* SP x 1.1 margin, A-M-188 margin class *)
  POLY_STOCKFT-01_ALARM_LO := 0.009000000000000001 ;

  (* FLOW control loop - set-point from the graph basis *)
  POLY_STOCKFT-02_SP := 0.0 ;  (* graph basis: STOCK_TO_FIBER normal 0.00 L/h )
  FB_PI_POLY_STOCKFT-02( PV := POLY_STOCKFT-02_PV, SP := POLY_STOCKFT-02_SP );  (* PI per AQS-CTL-002; GAIN/KI entered at commissioning from the step test (AQS-COM-001 sec. 3), anti-windup clamp per this FB *)
  POLY_STOCKFT-02_ALARM_HI := 0.0 ;  (* expected-zero state: any positive PV alarms )

  (* PRESSURE monitoring block - indication, no set-point invented )
  FB_AI_POLY_STOCKPT-01( PV := POLY_STOCKPT-01_PV );
  POLY_STOCKPT-01_ALARM_HI := 9.0 ;  (* 90 % of span, registered LSH convention )

  (* TEMPERATURE monitoring block - indication, no set-point invented )
  FB_AI_POLY_STOCKTE-01( PV := POLY_STOCKTE-01_PV );
  POLY_STOCKTE-01_ALARM_HI := 135.0 ;  (* 90 % of span, registered LSH convention )

  (* PRESSURE monitoring block - indication, no set-point invented )
  FB_AI_POWDER_RESINPT-01( PV := POWDER_RESINPT-01_PV );
  POWDER_RESINPT-01_ALARM_HI := 9.0 ;  (* 90 % of span, registered LSH convention )

  (* TEMPERATURE monitoring block - indication, no set-point invented )
  FB_AI_POWDER_RESINTE-01( PV := POWDER_RESINTE-01_PV );
  POWDER_RESINTE-01_ALARM_HI := 135.0 ;  (* 90 % of span, registered LSH convention )

  (* FLOW control loop - set-point from the graph basis *)
  TFE_SYNFT-01_SP := 0.0 ;  (* graph basis: TFE_TO_POLY_F normal 0.00 L/h )
  FB_PI_TFE_SYNFT-01( PV := TFE_SYNFT-01_PV, SP := TFE_SYNFT-01_SP );  (* PI per AQS-CTL-002; GAIN/KI entered at commissioning from the step test (AQS-COM-001 sec. 3), anti-windup clamp per this FB *)
  TFE_SYNFT-01_ALARM_HI := 0.0 ;  (* expected-zero state: any positive PV alarms )

  (* FLOW control loop - set-point from the graph basis *)
  TFE_SYNFT-02_SP := 0.01 ;  (* graph basis: TFE_HCL_TO_CRU normal 0.01 L/h )
  FB_PI_TFE_SYNFT-02( PV := TFE_SYNFT-02_PV, SP := TFE_SYNFT-02_SP );  (* PI per AQS-CTL-002; GAIN/KI entered at commissioning from the step test (AQS-COM-001 sec. 3), anti-windup clamp per this FB *)
  TFE_SYNFT-02_ALARM_HI := 0.011000000000000001 ;  (* SP x 1.1 margin, A-M-188 margin class *)
  TFE_SYNFT-02_ALARM_LO := 0.009000000000000001 ;

  (* LEVEL monitoring block - indication, no set-point invented )
  FB_AI_TFE_SYNLT-01( PV := TFE_SYNLT-01_PV );
  TFE_SYNLT-01_ALARM_HI := 90.0 ;  (* 90 % of span, registered LSH convention )

  (* PRESSURE monitoring block - indication, no set-point invented )
  FB_AI_TFE_SYNPT-01( PV := TFE_SYNPT-01_PV );
  TFE_SYNPT-01_ALARM_HI := 9.0 ;  (* 90 % of span, registered LSH convention )

  (* TEMPERATURE monitoring block - indication, no set-point invented )
  FB_AI_TFE_SYNTE-01( PV := TFE_SYNTE-01_PV );
  TFE_SYNTE-01_ALARM_HI := 135.0 ;  (* 90 % of span, registered LSH convention )

  (* FLOW control loop - set-point from the graph basis *)
  VDF_SYNFT-01_SP := 0.01 ;  (* graph basis: VDF_TO_POLY_F normal 0.01 L/h )
  FB_PI_VDF_SYNFT-01( PV := VDF_SYNFT-01_PV, SP := VDF_SYNFT-01_SP );  (* PI per AQS-CTL-002; GAIN/KI entered at commissioning from the step test (AQS-COM-001 sec. 3), anti-windup clamp per this FB *)
  VDF_SYNFT-01_ALARM_HI := 0.011000000000000001 ;  (* SP x 1.1 margin, A-M-188 margin class *)
  VDF_SYNFT-01_ALARM_LO := 0.009000000000000001 ;

  (* FLOW control loop - set-point from the graph basis *)
  VDF_SYNFT-02_SP := 0.02 ;  (* graph basis: VDF_HCL_TO_CRU normal 0.02 L/h )
  FB_PI_VDF_SYNFT-02( PV := VDF_SYNFT-02_PV, SP := VDF_SYNFT-02_SP );  (* PI per AQS-CTL-002; GAIN/KI entered at commissioning from the step test (AQS-COM-001 sec. 3), anti-windup clamp per this FB *)
  VDF_SYNFT-02_ALARM_HI := 0.022000000000000002 ;  (* SP x 1.1 margin, A-M-188 margin class *)
  VDF_SYNFT-02_ALARM_LO := 0.018000000000000002 ;

  (* LEVEL monitoring block - indication, no set-point invented )
  FB_AI_VDF_SYNLT-01( PV := VDF_SYNLT-01_PV );
  VDF_SYNLT-01_ALARM_HI := 90.0 ;  (* 90 % of span, registered LSH convention )

  (* PRESSURE monitoring block - indication, no set-point invented )
  FB_AI_VDF_SYNPT-01( PV := VDF_SYNPT-01_PV );
  VDF_SYNPT-01_ALARM_HI := 9.0 ;  (* 90 % of span, registered LSH convention )

  (* TEMPERATURE monitoring block - indication, no set-point invented )
  FB_AI_VDF_SYNTE-01( PV := VDF_SYNTE-01_PV );
  VDF_SYNTE-01_ALARM_HI := 135.0 ;  (* 90 % of span, registered LSH convention )

  (* FLOW control loop - set-point from the graph basis *)
  POLY_FIBERFT-01_SP := 0.0 ;  (* graph basis: FIBER_SCRAP normal 0.00 L/h )
  FB_PI_POLY_FIBERFT-01( PV := POLY_FIBERFT-01_PV, SP := POLY_FIBERFT-01_SP );  (* PI per AQS-CTL-002; GAIN/KI entered at commissioning from the step test (AQS-COM-001 sec. 3), anti-windup clamp per this FB *)
  POLY_FIBERFT-01_ALARM_HI := 0.0 ;  (* expected-zero state: any positive PV alarms )

  (* FLOW control loop - set-point from the graph basis *)
  POLY_FIBERFT-02_SP := 0.0 ;  (* graph basis: FLEECE_TO_MFG normal 0.00 L/h )
  FB_PI_POLY_FIBERFT-02( PV := POLY_FIBERFT-02_PV, SP := POLY_FIBERFT-02_SP );  (* PI per AQS-CTL-002; GAIN/KI entered at commissioning from the step test (AQS-COM-001 sec. 3), anti-windup clamp per this FB *)
  POLY_FIBERFT-02_ALARM_HI := 0.0 ;  (* expected-zero state: any positive PV alarms )

  (* PRESSURE monitoring block - indication, no set-point invented )
  FB_AI_POLY_FIBERPT-01( PV := POLY_FIBERPT-01_PV );
  POLY_FIBERPT-01_ALARM_HI := 9.0 ;  (* 90 % of span, registered LSH convention )

  (* TEMPERATURE monitoring block - indication, no set-point invented )
  FB_AI_POLY_FIBERTE-01( PV := POLY_FIBERTE-01_PV );
  POLY_FIBERTE-01_ALARM_HI := 135.0 ;  (* 90 % of span, registered LSH convention )

  (* LEVEL monitoring block - indication, no set-point invented )
  FB_AI_ACID_PLANTLT-01( PV := ACID_PLANTLT-01_PV );
  ACID_PLANTLT-01_ALARM_HI := 90.0 ;  (* 90 % of span, registered LSH convention )

  (* PRESSURE monitoring block - indication, no set-point invented )
  FB_AI_ACID_PLANTPT-01( PV := ACID_PLANTPT-01_PV );
  ACID_PLANTPT-01_ALARM_HI := 9.0 ;  (* 90 % of span, registered LSH convention )

  (* TEMPERATURE monitoring block - indication, no set-point invented )
  FB_AI_ACID_PLANTTE-01( PV := ACID_PLANTTE-01_PV );
  ACID_PLANTTE-01_ALARM_HI := 135.0 ;  (* 90 % of span, registered LSH convention )

  (* HF monitoring block - indication, no set-point invented )
  FB_AI_HF_GENAE-01( PV := HF_GENAE-01_PV );
  HF_GENAE-01_ALARM_HI := 9.0 ;  (* 90 % of span, registered LSH convention )

  (* LEVEL monitoring block - indication, no set-point invented )
  FB_AI_POLY_CONDLT-01( PV := POLY_CONDLT-01_PV );
  POLY_CONDLT-01_ALARM_HI := 90.0 ;  (* 90 % of span, registered LSH convention )

  (* SPEED monitoring block - indication, no set-point invented )
  FB_AI_POWDER_RESINST-01( PV := POWDER_RESINST-01_PV );
  POWDER_RESINST-01_ALARM_HI := 90.0 ;  (* 90 % of span, registered LSH convention )

  (* SPEED monitoring block - indication, no set-point invented )
  FB_AI_FILM_CASTST-01( PV := FILM_CASTST-01_PV );
  FILM_CASTST-01_ALARM_HI := 90.0 ;  (* 90 % of span, registered LSH convention )

  (* LEVEL monitoring block - indication, no set-point invented )
  FB_AI_POLY_STOCKLT-01( PV := POLY_STOCKLT-01_PV );
  POLY_STOCKLT-01_ALARM_HI := 90.0 ;  (* 90 % of span, registered LSH convention )

  (* TEMPERATURE monitoring block - indication, no set-point invented )
  FB_AI_POLY_FIBERTIR-01( PV := POLY_FIBERTIR-01_PV );
  POLY_FIBERTIR-01_ALARM_HI := 270.0 ;  (* 90 % of span, registered LSH convention )

  (* FLOW monitoring block - indication, no set-point invented )
  FB_AI_POLY_FIBERFIT-01( PV := POLY_FIBERFIT-01_PV );
  POLY_FIBERFIT-01_ALARM_HI := 1.8 ;  (* 90 % of span, registered LSH convention )

  (* SIF watch passthrough, no action in the basic program )
  SIF_WATCH_HF_GENTE-90 := HF_GENTE-90 ;  (* to safety CPU pair, AQS-CTL-003 )

  (* SIF watch passthrough, no action in the basic program )
  SIF_WATCH_POLY_OLEFINTE-90 := POLY_OLEFINTE-90 ;  (* to safety CPU pair, AQS-CTL-003 )

END_PROGRAM

(* ---- PLC-PUMPED_HYDRO.st ---- *)
(* AQS-CTL-004 X-CTL-04: control program source, generated by flow_graph/control/plc_programs.py *)
(* Basis: AQS-CTL-001 INSTRUMENT_INDEX.csv, AQS-CTL-002 control architecture, graph set-points. *)
(* PLC-PUMPED_HYDRO: CPU redundant pair; IO counts AI 2 AO 0 DI 4 DO 2 (modules per AQS-CTL-002, 16-channel, 20 % spare) *)
PROGRAM PLC_PUMPED_HYDRO_CTRL
VAR
  (* 100 ms cyclic task per AQS-CTL-002 *)
  HYDRO_SETPT-01_PV : REAL ;  (* no design pressure on the graph )
  HYDRO_SETTE-01_PV : REAL ;  (* band by service )
END_VAR

  (* PRESSURE monitoring block - indication, no set-point invented )
  FB_AI_HYDRO_SETPT-01( PV := HYDRO_SETPT-01_PV );
  HYDRO_SETPT-01_ALARM_HI := 9.0 ;  (* 90 % of span, registered LSH convention )

  (* TEMPERATURE monitoring block - indication, no set-point invented )
  FB_AI_HYDRO_SETTE-01( PV := HYDRO_SETTE-01_PV );
  HYDRO_SETTE-01_ALARM_HI := 135.0 ;  (* 90 % of span, registered LSH convention )

END_PROGRAM
